RoboDK station: Yuktii_Robotic_Car_Painting_Cell.rdk

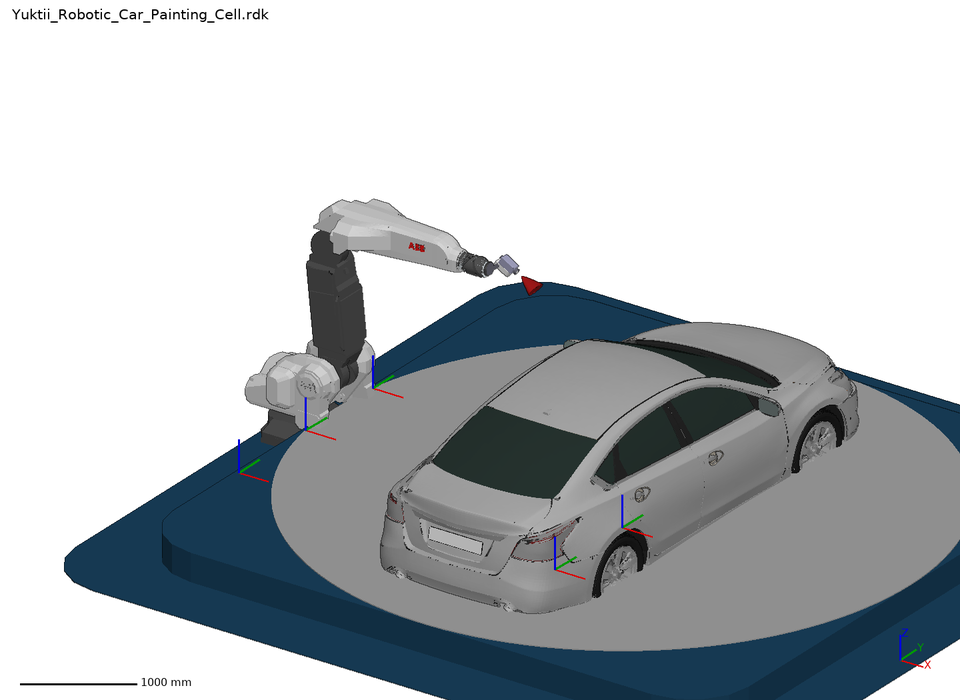
[picture v0: the station drawn from its stored meshes, robots at their saved joint values, targets as dots, program paths as lines]
Station Yuktii_Robotic_Car_Painting_Cell (saved by RoboDK 6.1.1). Poses are relative to the parent item; angles as X-Y-Z fixed-axis rotations.
  - frame ABB IRB 5400-22 Base at (0, 1000, 0) mm
    - robot ABB IRB 5400-22: 6 axes, payload 25 kg, reach 2829 mm, repeatability 0.15 mm, weight 1060 kg
        modified DH rows (alpha deg, a mm, theta deg, d mm): 0, 0, 0, 660; -90, 300, -90, 0; 0, 1200, 0, 0; -90, 213, -90, 1408.298; 35, 0, 0, 79.169; -70, 0, 180, 79.169
        base shift (0, 0, 0) mm, rotated rx 0 ry 0 rz 90 deg
        joint limits [-150, -65, -70, -720, -720, -720] to [150, 150, 70, 720, 720, 720]; home [0, 0, 0, 0, 0, 0]; saved at [-90, 0, 0, -0.001, 0.001, 0.001]
      - tool Generic Paint Sprayer, TCP at (50, 0, 450) mm, rotated rx 0 ry 30 rz 0 deg, size 277.6 x 203.2 x 501.7 mm
    - frame Painting Cell Frame at (0, 0, 0) mm
      - target Home (Cartesian target) at (2370, 0, 2023) mm, rotated rx -180 ry 60 rz -180 deg; joints [-90, 0, 0, 0, 0, 0] of ABB IRB 5400-22
        - target Home (Cartesian target) at (2370, 0, 2023) mm, rotated rx -180 ry 60 rz -180 deg; joints [-90, 0, 0, 0, 0, 0] of ABB IRB 5400-22
      - target Paint_Side_P01 (Cartesian target) at (2687.55, 277.64, 1440.42) mm, rotated rx -179.95 ry 58.29 rz -173.94 deg; joints [-85.31, 17.38, 3.62, 71.65, -55.76, -34.2] of ABB IRB 5400-22
      - target Paint_Side_P02 (Cartesian target) at (2657.17, 535.96, 1322.05) mm, rotated rx 179.9 ry 54.95 rz -168.86 deg; joints [-79.713, 18.918, 5.006, 71.33, -54.978, -34.463] of ABB IRB 5400-22
      - target Paint_Side_P03 (Cartesian target) at (2586.47, 830.84, 1163.47) mm, rotated rx 179.79 ry 50.46 rz -162.52 deg; joints [-73.303, 21.155, 6.646, 70.242, -53.863, -34.183] of ABB IRB 5400-22
      - target Paint_Side_P04 (Cartesian target) at (2523.64, 1053.32, 1068.21) mm, rotated rx 179.74 ry 48.21 rz -157.7 deg; joints [-68.45, 23.41, 6.64, 70.24, -53.86, -34.18] of ABB IRB 5400-22
      - target Paint_Side_P05 (Cartesian target) at (2478.28, 1238.02, 1045.31) mm, rotated rx 179.76 ry 48.45 rz -153.8 deg; joints [-64.55, 25.42, 4.99, 71.3, -54.96, -34.45] of ABB IRB 5400-22
      - target Paint_Side_P06 (Cartesian target) at (2451.93, 1495.48, 1004.92) mm, rotated rx 179.78 ry 49.69 rz -148.94 deg; joints [-59.68, 30.78, -0.3, 73.58, -57.34, -34.99] of ABB IRB 5400-22
      - target Paint_Side_P07 (Cartesian target) at (2459.02, 1865.41, 979.47) mm, rotated rx 179.83 ry 53.14 rz -143.1 deg; joints [-53.79, 41.5, -13.94, 74.57, -58.3, -35.26] of ABB IRB 5400-22
      - target Paint_Side_P08 (Cartesian target) at (2374.12, 1800.72, 860.49) mm, rotated rx 179.76 ry 48.46 rz -143.15 deg; joints [-53.84, 38.265, -5.941, 74.644, -58.451, -35.237] of ABB IRB 5400-22
      - target Paint_Side_P09 (Cartesian target) at (2351.62, 1976.72, 689.21) mm, rotated rx 179.72 ry 46.57 rz -140.3 deg; joints [-50.934, 45.88, -11.622, 74.742, -58.517, -35.278] of ABB IRB 5400-22
      - target Paint_Side_P10 (Cartesian target) at (2340.73, 2028.43, 516.1) mm, rotated rx 179.83 ry 43.58 rz -139.36 deg; joints [-48.072, 50.81, -13.693, -74.012, 58.304, 35.166] of ABB IRB 5400-22
      - target Paint_Side_P11 (Cartesian target) at (2319.85, 2100.8, 404.53) mm, rotated rx 176.79 ry 40.89 rz -141.32 deg; joints [-46.78, 54.89, -17.15, -68.32, 54.72, 34.95] of ABB IRB 5400-22
      - target Paint_Side_P12 (Cartesian target) at (2319.85, 2100.8, 404.53) mm, rotated rx 176.79 ry 40.89 rz -141.32 deg; joints [-48.695, 54.861, -16.957, 73.672, -54.894, -34.206] of ABB IRB 5400-22
      - target Paint_Side_P13 (Cartesian target) at (2357.01, 1967.98, 472.25) mm, rotated rx 176.8 ry 40.88 rz -143.6 deg; joints [-51.025, 50.456, -12.297, 74.028, -55.343, -34.246] of ABB IRB 5400-22
      - target Paint_Side_P14 (Cartesian target) at (2329.44, 1880.14, 669.1) mm, rotated rx 176.66 ry 43.13 rz -144.6 deg; joints [-52.014, 42.506, -6.735, 73.71, -55.102, -34.119] of ABB IRB 5400-22
      - target Paint_Side_P15 (Cartesian target) at (2356.38, 1841.89, 779.16) mm, rotated rx 176.49 ry 45.47 rz -145.61 deg; joints [-52.91, 40.16, -6.73, 73.71, -55.1, -34.11] of ABB IRB 5400-22
      - target Paint_Side_P16 (Cartesian target) at (2375.75, 1666.69, 808.98) mm, rotated rx 176.57 ry 44.12 rz -148.47 deg; joints [-55.911, 35.511, -1.417, 72.415, -53.828, -33.754] of ABB IRB 5400-22
      - target Paint_Side_P17 (Cartesian target) at (2358.71, 1489.22, 826.96) mm, rotated rx 176.71 ry 41.64 rz -151.09 deg; joints [-58.74, 30.11, 4.7, 69.11, -50.54, -32.85] of ABB IRB 5400-22
      - target Paint_Side_P18 (Cartesian target) at (2352.69, 1267.22, 769.5) mm, rotated rx 176.97 ry 36.54 rz -154.8 deg; joints [-62.721, 26.199, 10.485, 62.639, -44.318, -30.826] of ABB IRB 5400-22
      - target Paint_Side_P19 (Cartesian target) at (2339.07, 1164.01, 639.71) mm, rotated rx 177.2 ry 31.03 rz -156.46 deg; joints [-64.56, 26.76, 13.09, 57.4, -39.55, -28.91] of ABB IRB 5400-22
      - target Paint_Side_P20 (Cartesian target) at (2351.97, 1121.3, 477.66) mm, rotated rx 177.35 ry 27.01 rz -157.36 deg; joints [-65.53, 30.78, 13.09, 57.4, -39.55, -28.91] of ABB IRB 5400-22
      - target Paint_Side_P21 (Cartesian target) at (2354.18, 1035.31, 389.95) mm, rotated rx 111.95 ry -49.41 rz 97.65 deg; joints [-61.65, 33.04, 15.16, 173.91, -34.68, -354.54] of ABB IRB 5400-22
      - target Paint_Side_P22 (Cartesian target) at (2300.58, 869.96, 414.39) mm, rotated rx 111.93 ry -49.41 rz 94.75 deg; joints [-64.515, 28.088, 21.499, 170.665, -33.02, -351.904] of ABB IRB 5400-22
      - target Paint_Side_P23 (Cartesian target) at (2314.38, 611.77, 405.59) mm, rotated rx 112.89 ry -49.17 rz 88.15 deg; joints [-70.296, 25.908, 24.902, 169.511, -32.465, -350.855] of ABB IRB 5400-22
      - target Paint_Side_P24 (Cartesian target) at (2342.88, 284.67, 414.82) mm, rotated rx 112.88 ry -49.17 rz 80.3 deg; joints [-78.104, 24.346, 26.702, 169.017, -32.228, -350.379] of ABB IRB 5400-22
      - target Paint_Side_P25 (Cartesian target) at (2359.9, -36.58, 415.09) mm, rotated rx 112.87 ry -49.18 rz 72.49 deg; joints [-85.92, 24.34, 26.7, 169.01, -32.22, -350.37] of ABB IRB 5400-22
      - target Paint_Side_P26 (Cartesian target) at (2326.94, -394.75, 415.09) mm, rotated rx 112.87 ry -49.18 rz 63.75 deg; joints [-94.66, 24.34, 26.7, 169.01, -32.22, -350.37] of ABB IRB 5400-22
      - target Paint_Side_P27 (Cartesian target) at (2252.21, -705.72, 415.09) mm, rotated rx 112.87 ry -49.18 rz 55.98 deg; joints [-102.43, 24.34, 26.7, 169.01, -32.22, -350.37] of ABB IRB 5400-22
      - target Paint_Side_P28 (Cartesian target) at (2279.45, -959.44, 413.25) mm, rotated rx 112.85 ry -49.19 rz 50.17 deg; joints [-107.938, 28.675, 20.449, 174.163, -34.94, -354.053] of ABB IRB 5400-22
      - target Paint_Side_P29 (Cartesian target) at (2329.77, -987.72, 580.14) mm, rotated rx 106.08 ry -50.73 rz 55.16 deg; joints [-108.194, 26.054, 18.009, 175.068, -35.38, -354.858] of ABB IRB 5400-22
      - target Paint_Side_P30 (Cartesian target) at (2366.74, -1005.47, 624.94) mm, rotated rx 104.07 ry -51.08 rz 56.67 deg; joints [-108.306, 26.506, 15.801, 175.982, -35.848, -355.652] of ABB IRB 5400-22
      - target Paint_Side_P31 (Cartesian target) at (2341.49, -1086.77, 693.07) mm, rotated rx 101.34 ry -51.52 rz 56.91 deg; joints [-110.203, 25.189, 15.244, 176.226, -35.966, -355.862] of ABB IRB 5400-22
      - target Paint_Side_P32 (Cartesian target) at (2350.5, -1289.69, 809.61) mm, rotated rx 96.38 ry -52.11 rz 56.93 deg; joints [-114.207, 26.687, 9.223, 179.177, -37.505, -358.342] of ABB IRB 5400-22
      - target Paint_Side_P33 (Cartesian target) at (2338.83, -1380.36, 813.26) mm, rotated rx 96.14 ry -52.14 rz 55.32 deg; joints [-116.05, 28.1, 7.13, 180.3, -38.1, -359.26] of ABB IRB 5400-22
      - target Paint_Side_P34 (Cartesian target) at (2313.09, -1640.06, 805.87) mm, rotated rx 96.12 ry -52.15 rz 50.51 deg; joints [-120.978, 33.486, -0.37, 184.719, -40.559, -362.788] of ABB IRB 5400-22
      - target Paint_Side_P35 (Cartesian target) at (2385.33, -1800.15, 689.63) mm, rotated rx 99.75 ry -51.77 rz 45.91 deg; joints [-122.82, 42.83, -10.73, 191.42, -44.54, -367.93] of ABB IRB 5400-22
      - target Paint_Side_P36 (Cartesian target) at (2352.14, -1838.69, 532.96) mm, rotated rx 104.98 ry -51 rz 40.85 deg; joints [-123.79, 46.18, -10.73, 191.42, -44.54, -367.93] of ABB IRB 5400-22
      - target Paint_Side_P37 (Cartesian target) at (2383.84, -1926.08, 389.53) mm, rotated rx 109 ry -50.23 rz 36.81 deg; joints [-124.76, 53.4, -17.69, 196.12, -47.53, -371.4] of ABB IRB 5400-22
      - target Paint_Side_P38 (Cartesian target) at (2362.81, -2185.89, 442.85) mm, rotated rx 106.5 ry -50.73 rz 34.86 deg; joints [-128.68, 60.25, -31.28, 205.41, -53.93, -377.94] of ABB IRB 5400-22
      - target Paint_Side_P39 (Cartesian target) at (2368.83, -2190.72, 613.31) mm, rotated rx 101.33 ry -51.57 rz 38.89 deg; joints [-128.68, 56.9, -31.28, 205.41, -53.93, -377.94] of ABB IRB 5400-22
      - target Paint_Side_P40 (Cartesian target) at (2364.19, -2186.99, 852.08) mm, rotated rx 93.82 ry -52.34 rz 44.81 deg; joints [-128.68, 52.21, -31.28, 205.41, -53.93, -377.94] of ABB IRB 5400-22
      - target Paint_Side_P41 (Cartesian target) at (2429.25, -2245.53, 801.72) mm, rotated rx 95.27 ry -52.23 rz 43.67 deg; joints [-128.69, 58.91, -40.91, 211.91, -58.84, -382.23] of ABB IRB 5400-22
      - target Paint_Side_P42 (Cartesian target) at (2402.83, -2072.83, 809.3) mm, rotated rx 95.26 ry -52.24 rz 45.66 deg; joints [-126.674, 50.089, -26.385, 202.057, -51.536, -375.626] of ABB IRB 5400-22
      - target Paint_Side_P43 (Cartesian target) at (2397.72, -2068.76, 904.03) mm, rotated rx 92.18 ry -52.45 rz 48.11 deg; joints [-126.67, 48.19, -26.38, 202.05, -51.53, -375.62] of ABB IRB 5400-22
      - target Paint_Side_P44 (Cartesian target) at (2404.71, -1939.77, 930.5) mm, rotated rx 91.34 ry -52.5 rz 50.69 deg; joints [-124.73, 43.5, -19.74, 197.5, -48.43, -372.39] of ABB IRB 5400-22
      - target Paint_Side_P45 (Cartesian target) at (2424.76, -1763.9, 1025.75) mm, rotated rx 88.05 ry -52.62 rz 56.18 deg; joints [-121.803, 37.363, -13.341, 193.148, -45.618, -369.204] of ABB IRB 5400-22
      - target Paint_Side_P46 (Cartesian target) at (2501.66, -1816.71, 1075.26) mm, rotated rx 86.44 ry -52.65 rz 57.5 deg; joints [-121.814, 41.601, -21.433, 198.65, -49.191, -373.214] of ABB IRB 5400-22
      - target Paint_Side_P47 (Cartesian target) at (2521.68, -2035.45, 1120.54) mm, rotated rx 85.17 ry -52.65 rz 55.56 deg; joints [-124.802, 50.228, -36.673, 209.055, -56.613, -380.366] of ABB IRB 5400-22
      - target Paint_Side_P48 (Cartesian target) at (2491.9, -2224.63, 1126.16) mm, rotated rx 85.14 ry -52.65 rz 52.72 deg; joints [-127.67, 58.19, -50.18, 218.04, -63.79, -386.02] of ABB IRB 5400-22
      - target Paint_Side_P49 (Cartesian target) at (2637.88, -1982.32, 1160.05) mm, rotated rx 84.01 ry -52.64 rz 58.46 deg; joints [-122.825, 54.406, -44.865, 214.527, -60.901, -383.866] of ABB IRB 5400-22
      - target Paint_Side_P50 (Cartesian target) at (2582.23, -1809.13, 1242.07) mm, rotated rx 81.02 ry -52.57 rz 62.79 deg; joints [-120.85, 43.5, -29.72, 204.31, -53.12, -377.16] of ABB IRB 5400-22
      - target Paint_Side_P51 (Cartesian target) at (2618.31, -1589.81, 1315.52) mm, rotated rx 74.52 ry -52.89 rz 74.75 deg; joints [-117.93, 36.81, -20.97, 188.74, -39.61, -370.49] of ABB IRB 5400-22
      - target Paint_Side_P52 (Cartesian target) at (2623.91, -1459.92, 1331.56) mm, rotated rx 73.67 ry -52.77 rz 77.67 deg; joints [-115.766, 33.391, -16.372, 184.597, -37.067, -367.591] of ABB IRB 5400-22
      - target Paint_Side_P53 (Cartesian target) at (2616.77, -1306.34, 1411.32) mm, rotated rx 70.58 ry -52.28 rz 82.78 deg; joints [-113.193, 28.706, -12.08, 180.64, -34.713, -364.793] of ABB IRB 5400-22
      - target Paint_Side_P54 (Cartesian target) at (2683.21, -1167.98, 1441.11) mm, rotated rx 69.63 ry -52.12 rz 86.54 deg; joints [-110.175, 28.59, -12.841, 181.347, -35.125, -365.292] of ABB IRB 5400-22
      - target Paint_Side_P55 (Cartesian target) at (2649.23, -855.94, 1495.04) mm, rotated rx 66.81 ry -51.55 rz 94.56 deg; joints [-104.557, 21.072, -4.174, 173.152, -30.436, -359.425] of ABB IRB 5400-22
      - target Paint_Side_P56 (Cartesian target) at (2666.88, -565.19, 1525.15) mm, rotated rx 65.33 ry -51.24 rz 101.73 deg; joints [-98.61, 18.05, -1.14, 170.22, -28.81, -357.3] of ABB IRB 5400-22
      - target Paint_Side_P57 (Cartesian target) at (2662.07, -286.65, 1542.5) mm, rotated rx 64.33 ry -51 rz 108.4 deg; joints [-92.785, 15.593, 1.463, 167.684, -27.43, -355.464] of ABB IRB 5400-22
      - target Paint_Side_P58 (Cartesian target) at (2643.19, -58.71, 1533.21) mm, rotated rx 64.32 ry -51 rz 113.33 deg; joints [-87.918, 14.046, 3.678, 165.507, -26.262, -353.885] of ABB IRB 5400-22
      - target Paint_Side_P59 (Cartesian target) at (2643.6, 168.06, 1475.48) mm, rotated rx 66.28 ry -51.45 rz 116.71 deg; joints [-83.035, 14.713, 4.605, 164.582, -25.771, -353.214] of ABB IRB 5400-22
      - target Home (Cartesian target) at (2370, 0, 2023) mm, rotated rx -180 ry 60 rz 180 deg; joints [-90, 0, 0, -0.001, 0.001, 0] of ABB IRB 5400-22
      - target Target 64 (Cartesian target) at (2431.56, 1366.3, 1005.74) mm, rotated rx 179.72 ry 47.83 rz -151.03 deg; joints [-61.758, 26.931, 4.296, 71.642, -55.315, -34.517] of ABB IRB 5400-22
      - target Target 65 (Cartesian target) at (2421.45, 1107.77, 1017.39) mm, rotated rx 179.66 ry 44.84 rz -155.81 deg; joints [-66.537, 20.959, 10.51, 66.628, -50.22, -33.159] of ABB IRB 5400-22
      - target Target 66 (Cartesian target) at (2437.7, 946.12, 934.72) mm, rotated rx -171.38 ry 35.85 rz -163.72 deg; joints [-66.53, 20.95, 10.5, 66.62, -34.95, -48.93] of ABB IRB 5400-22
      - target Target 67 (Cartesian target) at (2455.17, 839.85, 965.83) mm, rotated rx -149.37 ry 33.2 rz -154.75 deg; joints [-66.53, 20.95, 10.5, 66.62, -34.95, -67.57] of ABB IRB 5400-22
      - target Target 68 (Cartesian target) at (2281.53, 854.15, 1189.47) mm, rotated rx -149.37 ry 33.21 rz -156.42 deg; joints [-63.59, 10.87, 13.54, 58.38, -21.49, -68.41] of ABB IRB 5400-22
      - target Target 69 (Cartesian target) at (2222.52, 748.18, 1108.21) mm, rotated rx -149.07 ry 23.15 rz -166.11 deg; joints [-63.59, 10.87, 13.54, 58.37, -6.99, -76.89] of ABB IRB 5400-22
      - target Target 70 (Cartesian target) at (2314.29, 671.58, 1031.07) mm, rotated rx -174.66 ry 26.9 rz 179.32 deg; joints [-69.41, 12.02, 14.02, 61.4, -11.65, -53.59] of ABB IRB 5400-22
      - target Target 71 (Cartesian target) at (2348.53, 655.22, 1084.89) mm, rotated rx -157.59 ry 30.49 rz -164.86 deg; joints [-69.41, 12.02, 14.02, 44.27, -11.65, -53.59] of ABB IRB 5400-22
      - target Target 72 (Cartesian target) at (2418.39, 483.96, 1040.28) mm, rotated rx -179 ry 31.42 rz 179.44 deg; joints [-76.21, 12.69, 14.02, 44.27, -11.65, -34.95] of ABB IRB 5400-22
      - target Target 73 (Cartesian target) at (2433.89, 322.66, 1024.16) mm, rotated rx -178.61 ry 30.12 rz 175.75 deg; joints [-79.63, 12.635, 13.993, 28.227, -0.687, -26.026] of ABB IRB 5400-22
      - target Target 74 (Cartesian target) at (2450.35, -154.11, 1024.41) mm, rotated rx -178.62 ry 30.13 rz 164.59 deg; joints [-90.78, 12.63, 13.99, 28.22, -0.68, -26.02] of ABB IRB 5400-22
      - target Target 75 (Cartesian target) at (2403.68, -533.92, 1101.06) mm, rotated rx -179.62 ry 33.41 rz 155.34 deg; joints [-100.12, 11.36, 13.92, 47.59, -14.17, -36.57] of ABB IRB 5400-22
      - target Target 76 (Cartesian target) at (2465.14, -650.21, 1055.69) mm, rotated rx -131.01 ry 24.44 rz -156.77 deg; joints [-103.4, 15.42, 13.83, 11.65, -26.09, -42.28] of ABB IRB 5400-22
      - target Target 77 (Cartesian target) at (2445.74, -924.66, 1070.36) mm, rotated rx -129.64 ry 26.09 rz -161.04 deg; joints [-109.805, 18.069, 10.791, 17.454, -31.485, -45.09] of ABB IRB 5400-22
      - target Target 78 (Cartesian target) at (2460.91, -1184.92, 1107) mm, rotated rx -127.19 ry 28.8 rz -163.21 deg; joints [-115.43, 22.74, 4.69, 23.29, -37.86, -47.32] of ABB IRB 5400-22
      - target Target 79 (Cartesian target) at (2442.56, -1519.43, 1130.02) mm, rotated rx -124.71 ry 31.02 rz -166.45 deg; joints [-122.1, 29.121, -3.711, 25.815, -41.925, -47.576] of ABB IRB 5400-22
      - target Target 80 (Cartesian target) at (2573.73, -1565.02, 1176.52) mm, rotated rx -122.14 ry 33.12 rz -163.1 deg; joints [-121.84, 35.09, -12.99, 25.26, -43.26, -46.09] of ABB IRB 5400-22
      - target Target 81 (Cartesian target) at (2490.66, -1694.09, 1176.52) mm, rotated rx -122.14 ry 33.12 rz -166.02 deg; joints [-124.76, 35.09, -12.99, 25.26, -43.26, -46.09] of ABB IRB 5400-22
      - target Target 82 (Cartesian target) at (2506.42, -1705.03, 1062.97) mm, rotated rx -124.25 ry 31.52 rz -167.15 deg; joints [-124.76, 37.48, -12.99, 25.26, -43.26, -46.09] of ABB IRB 5400-22
      - target Target 83 (Cartesian target) at (2447.26, -1788.9, 1062.97) mm, rotated rx -124.25 ry 31.52 rz -169.09 deg; joints [-126.7, 37.48, -12.99, 25.26, -43.26, -46.09] of ABB IRB 5400-22
      - target Target 84 (Cartesian target) at (2436.51, -1757.57, 963.26) mm, rotated rx -126.53 ry 29.7 rz -170.25 deg; joints [-126.265, 37.632, -10.258, 25.738, -43.152, -46.635] of ABB IRB 5400-22
      - target Target 85 (Cartesian target) at (2455.15, -1486.92, 1079.17) mm, rotated rx -108.62 ry 13.32 rz -151.02 deg; joints [-122.27, 29.83, -2.45, 6.99, -44.27, -53.59] of ABB IRB 5400-22
      - target Target 86 (Cartesian target) at (2383.23, -1251.24, 985.09) mm, rotated rx 137.84 ry 45.33 rz 149.2 deg; joints [-127.093, 29.212, 4.635, 62.346, -71.879, 16.542] of ABB IRB 5400-22
      - target Target 87 (Cartesian target) at (2389.27, -903.36, 973.08) mm, rotated rx 136.67 ry 40.82 rz 160.1 deg; joints [-121.56, 24.75, 9.87, 54.4, -70.28, 23.75] of ABB IRB 5400-22
      - target Target 88 (Cartesian target) at (2356.03, -724.5, 1025.32) mm, rotated rx 136.02 ry 38.81 rz 167.16 deg; joints [-119.008, 21.071, 11.864, 47.567, -68.887, 30.048] of ABB IRB 5400-22
      - target Target 89 (Cartesian target) at (2379.15, -397.54, 973.43) mm, rotated rx 134.16 ry 33.87 rz 178.02 deg; joints [-112.26, 21.4, 12.24, 40.3, -67.78, 37.13] of ABB IRB 5400-22
      - target Target 90 (Cartesian target) at (2365.39, -354.45, 922.39) mm, rotated rx 132.55 ry 30.09 rz -178.82 deg; joints [-111.726, 22.838, 11.574, 35.485, -67.33, 42.068] of ABB IRB 5400-22
      - target Target 91 (Cartesian target) at (2377.11, -152.88, 925.3) mm, rotated rx 132.01 ry 28.94 rz -172.71 deg; joints [-107.078, 22.996, 10.964, 33.204, -67.266, 44.598] of ABB IRB 5400-22
      - target Target 93 (Cartesian target) at (2365.62, 454.26, 908.58) mm, rotated rx -180 ry 29.04 rz -169.13 deg; joints [-79.13, 12.02, 18.94, 0, 0, 0] of ABB IRB 5400-22
      - target Target 93 (Cartesian target) at (2307.39, 692.25, 908.9) mm, rotated rx -180 ry 29.05 rz -163.3 deg; joints [-73.3, 12.02, 18.93, 0, 0, 0] of ABB IRB 5400-22
      - target Target 94 (Cartesian target) at (2321.31, 696.8, 661.14) mm, rotated rx 179.99 ry 22.35 rz -163.31 deg; joints [-73.29, 18.72, 18.93, -0.01, 0.02, 0.01] of ABB IRB 5400-22
      - target Target 96 (Cartesian target) at (2265.55, 985.02, 820.27) mm, rotated rx 179.99 ry 29.71 rz -156.52 deg; joints [-65.754, 16.526, 17.771, -34.157, 22.81, 19.698] of ABB IRB 5400-22
      - target Target 96 (Cartesian target) at (2355.77, 1024.1, 856.74) mm, rotated rx 179.89 ry 35.33 rz -156.57 deg; joints [-65.504, 19.848, 14.513, -52.037, 36.976, 28.267] of ABB IRB 5400-22
      - target Target 97 (Cartesian target) at (2297.33, 1237.75, 742.18) mm, rotated rx 179.94 ry 33.8 rz -151.73 deg; joints [-60.656, 24.16, 13.203, -55.596, 40.098, 29.701] of ABB IRB 5400-22
      - target Target 99 (Cartesian target) at (2334.09, -1564.72, 911.12) mm, rotated rx 179.66 ry 44.54 rz 145.94 deg; joints [-122.78, 29.44, 3.24, -68.04, 51.94, 33.9] of ABB IRB 5400-22
      - target Target 99 (Cartesian target) at (2383.08, -1922.61, 792.43) mm, rotated rx 129.8 ry 40.18 rz 114.6 deg; joints [-131.6, 45.51, -12.13, -71.68, 58.25, 72.23] of ABB IRB 5400-22
      - target Target 100 (Cartesian target) at (2320.47, -1611.26, 821.25) mm, rotated rx 131.5 ry 37.1 rz 123.46 deg; joints [-128.622, 34.639, 2.593, -77.933, 59.044, 77.036] of ABB IRB 5400-22
      - target Target 101 (Cartesian target) at (2345.57, -1090.33, 826.64) mm, rotated rx 133.32 ry 31.79 rz 139.56 deg; joints [-120.514, 24.999, 14.295, -81.52, 53.807, 82.959] of ABB IRB 5400-22
      - target Target 102 (Cartesian target) at (2357.6, -322.96, 677.83) mm, rotated rx 134.67 ry 19.27 rz 165.08 deg; joints [-105.77, 21.651, 21.251, -84.321, 41.712, 92.046] of ABB IRB 5400-22
      - target Target 103 (Cartesian target) at (2336.63, 1100.19, 539.42) mm, rotated rx -169.54 ry 29.49 rz -173.27 deg; joints [-57.41, 31.45, 10.05, -33.99, 55.09, -1.39] of ABB IRB 5400-22
      - target Target 104 (Cartesian target) at (2301.03, -953.45, 610.69) mm, rotated rx 143.59 ry 28.63 rz 126.15 deg; joints [-112.14, 23.41, 22.34, -54.77, 58.25, 53.59] of ABB IRB 5400-22
      - target Target 105 (Cartesian target) at (2332.17, -895.94, 508.39) mm, rotated rx 131.34 ry 21.29 rz 122.4 deg; joints [-112.14, 27.43, 22.34, -54.77, 58.24, 67.57] of ABB IRB 5400-22
      - target Target 106 (Cartesian target) at (2329.78, 1096.4, 434.09) mm, rotated rx -168.24 ry 27.08 rz -172.64 deg; joints [-57.4, 34.13, 10.04, -33.99, 55.09, -1.38] of ABB IRB 5400-22
      - target Home (Cartesian target) at (2370, 0, 2023) mm, rotated rx -180 ry 60 rz -180 deg; joints [-90, 0, 0, 0, 0, 0] of ABB IRB 5400-22
      - target New_Side1 (Cartesian target) at (2658.8, 275.75, 1524.52) mm, rotated rx -179.85 ry 60.31 rz -173.84 deg; joints [-85.3, 15.37, 3.61, 71.65, -55.76, -34.2] of ABB IRB 5400-22
      - target Target 108 (Cartesian target) at (2664.22, 523.99, 1523.09) mm, rotated rx -179.82 ry 60.98 rz -168.61 deg; joints [-80.075, 17.43, 1.429, 72.616, -56.756, -34.445] of ABB IRB 5400-22
      - target Target 109 (Cartesian target) at (2665.93, 762.89, 1510.03) mm, rotated rx -179.81 ry 61.52 rz -163.77 deg; joints [-75.205, 20.33, -1.486, 73.532, -57.694, -34.668] of ABB IRB 5400-22
      - target Target 110 (Cartesian target) at (2659.82, 1167.43, 1438.23) mm, rotated rx -179.83 ry 61.51 rz -156.05 deg; joints [-67.415, 27.34, -7.983, 74.44, -58.603, -34.91] of ABB IRB 5400-22
      - target Target 111 (Cartesian target) at (2634.53, 1372.82, 1374.32) mm, rotated rx -179.9 ry 60.79 rz -152.28 deg; joints [-63.559, 31.151, -11.105, 74.432, -58.556, -34.922] of ABB IRB 5400-22
      - target Target 112 (Cartesian target) at (2613.56, 1565.5, 1326.63) mm, rotated rx -156.73 ry 55.5 rz -141.8 deg; joints [-57.009, 36.126, -17.739, 72.955, -48.745, -56.751] of ABB IRB 5400-22
      - target Target 113 (Cartesian target) at (2569.84, 1720.18, 1273.47) mm, rotated rx -156.83 ry 54.94 rz -138.73 deg; joints [-54.23, 38.988, -20.195, 72.171, -48.363, -56.199] of ABB IRB 5400-22
      - target Target 114 (Cartesian target) at (2584.39, 1876.48, 1194.72) mm, rotated rx -130.83 ry 49.71 rz -130.74 deg; joints [-48.997, 49.602, -32.053, 80.685, -47.963, -85.459] of ABB IRB 5400-22
      - target Target 115 (Cartesian target) at (2561.17, 2039.05, 1143.93) mm, rotated rx -130.84 ry 49.71 rz -126.9 deg; joints [-46.823, 54.832, -38.834, 75.333, -44.25, -82.66] of ABB IRB 5400-22
      - target Target 116 (Cartesian target) at (2560.42, 2235.82, 1117.58) mm, rotated rx -130.52 ry 50.72 rz -122.04 deg; joints [-44.699, 64.532, -54.336, 60.957, -33.248, -75.821] of ABB IRB 5400-22
      - target Target 117 (Cartesian target) at (2472.08, 1830.68, 1089.48) mm, rotated rx -131.27 ry 45.32 rz -133.48 deg; joints [-47.68, 44.84, -21.46, 88.72, -52.51, -90.54] of ABB IRB 5400-22
      - target Target 118 (Cartesian target) at (2481.64, 1840.12, 992.4) mm, rotated rx -131.47 ry 43.32 rz -133.61 deg; joints [-47.67, 46.85, -21.46, 88.72, -52.51, -90.54] of ABB IRB 5400-22
      - target Target 119 (Cartesian target) at (2403.75, 1952.84, 974.82) mm, rotated rx -131.49 ry 43.1 rz -131.1 deg; joints [-45.15, 47.52, -21.91, 88.72, -52.51, -90.54] of ABB IRB 5400-22
      - target Target 120 (Cartesian target) at (2386.21, 2042.31, 939.94) mm, rotated rx -118.24 ry 38.52 rz -123.55 deg; joints [-43.2, 52.21, -26.67, 84.98, -50.64, -100.19] of ABB IRB 5400-22
      - target Target 121 (Cartesian target) at (2451.41, 2090.3, 884.4) mm, rotated rx -118.24 ry 38.52 rz -121.61 deg; joints [-43.82, 57.066, -32.806, 78.784, -47.107, -96.687] of ABB IRB 5400-22
      - target Target 122 (Cartesian target) at (2455.32, 2094.41, 790.53) mm, rotated rx -118.74 ry 36.71 rz -121.91 deg; joints [-43.82, 58.91, -32.8, 78.78, -47.1, -96.68] of ABB IRB 5400-22
      - target Target 123 (Cartesian target) at (2455.32, 2094.41, 790.53) mm, rotated rx -118.74 ry 36.71 rz -121.91 deg; joints [-43.82, 58.91, -32.8, 78.78, -47.1, -96.68] of ABB IRB 5400-22
      - target Target 124 (Cartesian target) at (2404.28, 2248.71, 785.39) mm, rotated rx -105.86 ry 31.76 rz -113.98 deg; joints [-40.99, 65.21, -41.48, 70.02, -41.43, -104.85] of ABB IRB 5400-22
      - target Target 125 (Cartesian target) at (2471.68, 2333.46, 771.99) mm, rotated rx -105.61 ry 32.35 rz -110.71 deg; joints [-41.26, 72.98, -55.01, 51.48, -28.89, -95.09] of ABB IRB 5400-22
      - target Target 126 (Cartesian target) at (2420.97, 2346.66, 641.9) mm, rotated rx -106.69 ry 29.85 rz -111.27 deg; joints [-40.388, 73.008, -50.637, 57.956, -33.304, -98.515] of ABB IRB 5400-22
      - target Target 127 (Cartesian target) at (2419.04, 2345.11, 536.48) mm, rotated rx -107.43 ry 27.97 rz -111.62 deg; joints [-40.38, 74.98, -50.63, 57.95, -33.3, -98.51] of ABB IRB 5400-22
      - target Target 128 (Cartesian target) at (2416.56, 2342.24, 464.73) mm, rotated rx -107.92 ry 26.7 rz -111.84 deg; joints [-40.38, 76.32, -50.62, 57.95, -33.3, -98.5] of ABB IRB 5400-22
      - target Target 129 (Cartesian target) at (2372.36, 2151.25, 436.56) mm, rotated rx -108.49 ry 24.41 rz -118.69 deg; joints [-41.3, 67.62, -33.69, 79.97, -47.44, -109.64] of ABB IRB 5400-22
      - target Target 130 (Cartesian target) at (2332.85, 1868.98, 420.57) mm, rotated rx -108.74 ry 20.64 rz -131.35 deg; joints [-42.87, 60.25, -19.97, 102.16, -57.85, -121.49] of ABB IRB 5400-22
      - target Target 131 (Cartesian target) at (2362.92, 1786.92, 599.14) mm, rotated rx -108.64 ry 23.66 rz -135.23 deg; joints [-44.065, 55.5, -18.473, 106.546, -59.354, -124.195] of ABB IRB 5400-22
      - target Target 132 (Cartesian target) at (2352.74, 1670.01, 745.54) mm, rotated rx -108.35 ry 24.36 rz -143.99 deg; joints [-44.63, 51.54, -17.35, 119.07, -63.26, -132.98] of ABB IRB 5400-22
      - target Target 133 (Cartesian target) at (2352.74, 1670.01, 745.54) mm, rotated rx -108.35 ry 24.36 rz -143.99 deg; joints [-44.63, 51.54, -17.35, 119.07, -63.26, -132.98] of ABB IRB 5400-22
      - target Target 134 (Cartesian target) at (2336.83, 1664.58, 784.26) mm, rotated rx -108.35 ry 24.36 rz -146.45 deg; joints [-44.2, 51.085, -18.114, 123.264, -64.411, -136.171] of ABB IRB 5400-22
      - target Target 135 (Cartesian target) at (2327.68, 1352.65, 832.3) mm, rotated rx -103.03 ry 1.48 rz -109.02 deg; joints [-54.222, 28.746, 9.244, -28.437, 5.83, -416.904] of ABB IRB 5400-22
      - target Target 136 (Cartesian target) at (2306.29, 1190.11, 834.99) mm, rotated rx -103.59 ry 0.51 rz -109.04 deg; joints [-57.25, 24.08, 15.62, -46.54, 14.38, -405.66] of ABB IRB 5400-22
      - target Target 137 (Cartesian target) at (2334.57, 1071.93, 714.75) mm, rotated rx -105.67 ry -2.13 rz -112.44 deg; joints [-59.663, 25.899, 17.118, -42.65, 12.894, -408.122] of ABB IRB 5400-22
      - target Target 138 (Cartesian target) at (2330.83, 977.71, 595.32) mm, rotated rx -107.81 ry -4.94 rz -115.26 deg; joints [-61.28, 27.482, 18.954, -36.885, 10.544, -411.674] of ABB IRB 5400-22
      - target Target 174 (Cartesian target) at (2370, 0, 2023) mm, rotated rx -180 ry 60 rz -180 deg; joints [-90, 0, 0, 0, 0, 0] of ABB IRB 5400-22
      - target Target 175 (Cartesian target) at (2003.56, 0, 1478.8) mm, rotated rx -180 ry 46.35 rz -180 deg; joints [-90, -16.78, 30.43, 0, 0, 0] of ABB IRB 5400-22
      - target Target 140 (Cartesian target) at (2346.95, 903.39, 372.64) mm, rotated rx 105.05 ry -53.98 rz 91.43 deg; joints [-62.798, 32.643, 18.247, 171.995, -33.643, 20.163] of ABB IRB 5400-22
      - target Target 141 (Cartesian target) at (2342.97, 174.12, 368.94) mm, rotated rx 106.29 ry -53.62 rz 73.14 deg; joints [-79.038, 26.889, 26.977, 168.799, -32.261, 24.129] of ABB IRB 5400-22
      - target Target 142 (Cartesian target) at (2350.11, -835.78, 365.76) mm, rotated rx 105.46 ry -53.86 rz 50.44 deg; joints [-103.37, 32.12, 19.32, 171.49, -33.41, 20.69] of ABB IRB 5400-22
      - target Target 143 (Cartesian target) at (2337.88, -1111.77, 373.69) mm, rotated rx 100.3 ry -27.32 rz 78.87 deg; joints [-114.08, 34.8, 19.32, 123.5, -33.41, 25.63] of ABB IRB 5400-22
      - target Target 145 (Cartesian target) at (2293.54, -1236.73, 723.48) mm, rotated rx 90.92 ry -25.06 rz 80.1 deg; joints [-116.99, 26.09, 19.32, 123.5, -33.41, 25.63] of ABB IRB 5400-22
      - target Target 146 (Cartesian target) at (2289.45, -1364.49, 777.87) mm, rotated rx 89.51 ry -24.66 rz 77.78 deg; joints [-119.341, 27.215, 15.821, 125.411, -33.698, 23.861] of ABB IRB 5400-22
      - target Target 147 (Cartesian target) at (2331.68, -1489.87, 827.19) mm, rotated rx 88.33 ry -24.33 rz 75.77 deg; joints [-120.96, 30.317, 9.647, 128.755, -34.187, 20.613] of ABB IRB 5400-22
      - target Target 148 (Cartesian target) at (2325.53, -1697.75, 857.4) mm, rotated rx 90.71 ry -12.89 rz 74.04 deg; joints [-124.76, 34.8, 3.22, 131.19, -44.16, 13.4] of ABB IRB 5400-22
      - target Target 149 (Cartesian target) at (2344.83, -1796.94, 780.88) mm, rotated rx 92.31 ry -13.4 rz 71.83 deg; joints [-125.99, 39.49, -1.41, 132.9, -44.03, 11.23] of ABB IRB 5400-22
      - target Target 150 (Cartesian target) at (2326.9, -1929.07, 663.98) mm, rotated rx 94.68 ry -14.1 rz 68.63 deg; joints [-128.1, 44.84, -5.96, 134.54, -43.87, 9.06] of ABB IRB 5400-22
      - target Target 151 (Cartesian target) at (2330.1, -2009.3, 463.73) mm, rotated rx 98.67 ry -15.23 rz 66.11 deg; joints [-129.136, 51.704, -10.429, 136.139, -43.668, 6.9] of ABB IRB 5400-22
      - target Target 152 (Cartesian target) at (2324.17, -2004.03, 374.06) mm, rotated rx 100.53 ry -15.71 rz 65.62 deg; joints [-129.13, 53.55, -10.42, 136.13, -43.66, 6.9] of ABB IRB 5400-22
      - target Target 153 (Cartesian target) at (2350.91, -2138.26, 409.75) mm, rotated rx 95.5 ry -11.04 rz 69.58 deg; joints [-131.63, 58.24, -17.66, 125.27, -42.28, 12.86] of ABB IRB 5400-22
      - target Target 154 (Cartesian target) at (2358.16, -2144.71, 578.33) mm, rotated rx 92.34 ry -9.81 rz 70.15 deg; joints [-131.63, 54.89, -17.66, 125.27, -42.28, 12.86] of ABB IRB 5400-22
      - target Target 155 (Cartesian target) at (2351.78, -2034.83, 598.74) mm, rotated rx 92.01 ry -9.71 rz 72.24 deg; joints [-130.35, 50.87, -11.47, 123.69, -43.37, 15.86] of ABB IRB 5400-22
      - target Target 156 (Cartesian target) at (2361.73, -2031.04, 641.31) mm, rotated rx 91.21 ry -9.37 rz 72.51 deg; joints [-130.17, 50.2, -11.81, 123.77, -43.3, 15.68] of ABB IRB 5400-22
      - target Target 157 (Cartesian target) at (2381.46, -2007.86, 641.31) mm, rotated rx 91.21 ry -9.37 rz 73.07 deg; joints [-129.61, 50.2, -11.81, 123.77, -43.3, 15.68] of ABB IRB 5400-22
      - target Target 158 (Cartesian target) at (2371.55, -1954.82, 707.1) mm, rotated rx 89.96 ry -8.85 rz 74.24 deg; joints [-129.052, 47.01, -8.72, 122.993, -43.864, 17.153] of ABB IRB 5400-22
      - target Target 159 (Cartesian target) at (2375.07, -1837.16, 777.79) mm, rotated rx 88.57 ry -8.25 rz 76.8 deg; joints [-127.418, 42.553, -3.828, 121.744, -44.753, 19.458] of ABB IRB 5400-22
      - target Target 160 (Cartesian target) at (2381.93, -1755.68, 825.25) mm, rotated rx 87.62 ry -7.82 rz 78.62 deg; joints [-126.181, 39.789, -1.019, 121.01, -45.257, 20.759] of ABB IRB 5400-22
      - target Target 161 (Cartesian target) at (2414.53, -1737.26, 915.15) mm, rotated rx 85.9 ry -7.01 rz 79.3 deg; joints [-125.47, 38.82, -2.55, 121.42, -44.98, 20.01] of ABB IRB 5400-22
      - target Target 162 (Cartesian target) at (2430.75, -1523.5, 926.8) mm, rotated rx 85.49 ry -6.84 rz 83.96 deg; joints [-122.07, 34.13, 4.33, 119.51, -46.13, 23.25] of ABB IRB 5400-22
      - target Target 163 (Cartesian target) at (2440.67, -1339.39, 956.51) mm, rotated rx 84.74 ry -6.46 rz 88.16 deg; joints [-118.98, 30.11, 9.37, 118.02, -46.96, 25.58] of ABB IRB 5400-22
      - target Target 164 (Cartesian target) at (2475.14, -1166.95, 1009.48) mm, rotated rx 83.54 ry -5.85 rz 92.22 deg; joints [-115.594, 27.22, 11.797, 117.241, -47.321, 26.717] of ABB IRB 5400-22
      - target Target 165 (Cartesian target) at (2541.7, -966.33, 1114.32) mm, rotated rx 81.35 ry -4.68 rz 96.85 deg; joints [-111.17, 24.75, 11.79, 117.24, -47.32, 26.71] of ABB IRB 5400-22
      - target Target 166 (Cartesian target) at (2438.77, -1046.57, 1116.61) mm, rotated rx 127.47 ry 31.35 rz 100.95 deg; joints [-111.17, 19.39, 11.78, 123.5, -62.91, -30.29] of ABB IRB 5400-22
      - target Target 167 (Cartesian target) at (2502.55, -919.8, 1181.69) mm, rotated rx 125.46 ry 32.41 rz 102.81 deg; joints [-108.097, 19.012, 10.424, 123.971, -63.426, -30.24] of ABB IRB 5400-22
      - target Target 168 (Cartesian target) at (2593.39, -572.94, 1327.96) mm, rotated rx 121.36 ry 34.36 rz 108.17 deg; joints [-100.33, 16.71, 9.02, 124.4, -63.89, -30.21] of ABB IRB 5400-22
      - target Target 169 (Cartesian target) at (2593.39, -572.94, 1327.96) mm, rotated rx 121.36 ry 34.36 rz 108.17 deg; joints [-100.33, 16.71, 9.02, 124.4, -63.89, -30.21] of ABB IRB 5400-22
      - target Target 170 (Cartesian target) at (2606.86, -356.08, 1410.12) mm, rotated rx 119.19 ry 35.3 rz 111.63 deg; joints [-95.63, 14.7, 9.02, 124.4, -63.89, -30.21] of ABB IRB 5400-22
      - target Target 171 (Cartesian target) at (2660.01, 12.46, 1498.43) mm, rotated rx 116.04 ry 36.56 rz 117.57 deg; joints [-87.53, 15.37, 5.88, 125.22, -64.73, -30.24] of ABB IRB 5400-22
      - target Target 172 (Cartesian target) at (2657.4, 365.18, 1513.99) mm, rotated rx 115.28 ry 36.85 rz 124.54 deg; joints [-79.958, 16.341, 4.355, 125.548, -65.04, -30.288] of ABB IRB 5400-22
      - target Home (Cartesian target) at (2370, 0, 2023) mm, rotated rx -180 ry 60 rz -180 deg; joints [-90, 0, 0, 0, 0, 0] of ABB IRB 5400-22
      - target Target 175 (Cartesian target) at (2472.08, 1830.68, 1089.48) mm, rotated rx -131.27 ry 45.32 rz -133.48 deg; joints [-47.68, 44.84, -21.46, 88.72, -52.51, -90.54] of ABB IRB 5400-22
      - target Target 176 (Cartesian target) at (2427.86, 1264.35, 1099.18) mm, rotated rx -130.5 ry 36.23 rz -154.16 deg; joints [-53.543, 32.02, -4.416, 109.606, -56.215, -109.469] of ABB IRB 5400-22
      - target Target 177 (Cartesian target) at (2382.88, -673.82, 1025.37) mm, rotated rx -179.04 ry 31.47 rz 152.37 deg; joints [-103.4, 13.36, 13.92, 47.58, -14.16, -36.56] of ABB IRB 5400-22
      - target Target 178 (Cartesian target) at (2295.9, -645.43, 1322.87) mm, rotated rx 178.75 ry 38.01 rz 151.12 deg; joints [-102.66, 4.66, 13.84, 21.49, 3.52, -21.94] of ABB IRB 5400-22
      - target Target 179 (Cartesian target) at (2289.84, -801.89, 1175.32) mm, rotated rx -179.9 ry 34.14 rz 148.27 deg; joints [-106.31, 8.68, 13.84, 21.49, 3.52, -21.94] of ABB IRB 5400-22
      - target Target 180 (Cartesian target) at (2275.94, -840.54, 1175.32) mm, rotated rx -179.9 ry 34.14 rz 147.3 deg; joints [-107.28, 8.68, 13.84, 21.49, 3.52, -21.94] of ABB IRB 5400-22
      - target Target 181 (Cartesian target) at (2192.36, -786.89, 1107.97) mm, rotated rx -179.9 ry 34.14 rz 147.3 deg; joints [-105.797, 5.265, 20.224, -4.848, 20.771, -6.041] of ABB IRB 5400-22
      - target Target 182 (Cartesian target) at (2382.86, -994.11, 973.37) mm, rotated rx 178.01 ry 39.71 rz 144.57 deg; joints [-108.817, 18.689, 12.609, -41.483, 44.688, 16.144] of ABB IRB 5400-22
      - target Target 183 (Cartesian target) at (2400.81, -1006.99, 991.61) mm, rotated rx 177.52 ry 40.97 rz 144.26 deg; joints [-108.962, 19.291, 11.631, -43.669, 46.321, 17.307] of ABB IRB 5400-22
      - target Target 184 (Cartesian target) at (2376.37, -1347.22, 1008.7) mm, rotated rx 145.79 ry 38.45 rz 130.25 deg; joints [-121.27, 24.75, 5.8, -54.81, 42.93, 54.56] of ABB IRB 5400-22
      - target Target 185 (Cartesian target) at (2422.65, -1754.66, 920.86) mm, rotated rx 128.56 ry 37.29 rz 115.93 deg; joints [-128.64, 39.35, -8.65, -60.74, 49.18, 70.09] of ABB IRB 5400-22
      - target Target 186 (Cartesian target) at (2354.37, -1824.66, 835.51) mm, rotated rx 129.7 ry 35.34 rz 115.04 deg; joints [-130.58, 40.29, -7.39, -61.24, 49.21, 70.51] of ABB IRB 5400-22
      - target Target 187 (Cartesian target) at (2377.86, -1153.27, 879.75) mm, rotated rx 132.19 ry 29.42 rz 134.82 deg; joints [-120.75, 25.42, 10.41, -65.41, 42.63, 77.65] of ABB IRB 5400-22
      - target Target 188 (Cartesian target) at (2359.94, -929.24, 826.9) mm, rotated rx 133.34 ry 24.54 rz 142.99 deg; joints [-117.419, 22.585, 14.742, -64.911, 36.511, 80.455] of ABB IRB 5400-22
      - target Target 189 (Cartesian target) at (2391.23, -667.17, 827.39) mm, rotated rx 133.65 ry 22.34 rz 150.99 deg; joints [-112.14, 20.73, 16.41, -64.25, 32.39, 82.07] of ABB IRB 5400-22
      - target Target 190 (Cartesian target) at (2202.62, -831.48, 1034.88) mm, rotated rx 133.65 ry 22.34 rz 150.99 deg; joints [-118.843, 12.15, 18.199, -62.412, 21.357, 86.632] of ABB IRB 5400-22
      - target Target 191 (Cartesian target) at (2109.76, -912.38, 1137.03) mm, rotated rx 133.65 ry 22.34 rz 150.99 deg; joints [-122.36, 8.718, 17.956, -62.764, 16.398, 90.091] of ABB IRB 5400-22
      - target Target 192 (Cartesian target) at (2280.41, -644.54, 1108.05) mm, rotated rx 155.69 ry 31.8 rz 164.39 deg; joints [-111.17, 8.68, 17.95, -58.25, 20.97, 62.91] of ABB IRB 5400-22
      - target Target 193 (Cartesian target) at (2291.01, -605.37, 1108.38) mm, rotated rx 155.69 ry 31.81 rz 165.37 deg; joints [-110.19, 8.67, 17.95, -58.24, 20.96, 62.91] of ABB IRB 5400-22
      - target Target 194 (Cartesian target) at (2368.73, -670.39, 889.33) mm, rotated rx -161.9 ry 27.55 rz -170.95 deg; joints [-106.31, 14.7, 17.95, -67.57, 25.63, 30.29] of ABB IRB 5400-22
      - target Target 195 (Cartesian target) at (2390.69, -115.75, 865.83) mm, rotated rx -164.07 ry 23.28 rz -159.26 deg; joints [-93.654, 12.603, 19.045, -35.861, 2.338, 14.58] of ABB IRB 5400-22
      - target Target 196 (Cartesian target) at (2355.61, 340.8, 891.86) mm, rotated rx 176.44 ry 30.26 rz 172.94 deg; joints [-78.181, 11.623, 20.691, -16.162, 28.516, 5.142] of ABB IRB 5400-22
      - target Target 197 (Cartesian target) at (2340.91, 486.87, 938.41) mm, rotated rx -175.27 ry 39.05 rz 171.84 deg; joints [-70.439, 13.268, 20.61, -39.821, 58.372, 2.503] of ABB IRB 5400-22
      - target Target 198 (Cartesian target) at (2390.18, 1030.97, 973.44) mm, rotated rx -175.27 ry 39.05 rz 171.84 deg; joints [-57.416, 24.788, 4.133, -31.939, 65.368, -10.181] of ABB IRB 5400-22
      - target Target 199 (Cartesian target) at (2421.98, 1792.86, 985.86) mm, rotated rx -173.33 ry 37.83 rz 173.05 deg; joints [-44.166, 50.231, -35.31, -18.806, 69, -32.901] of ABB IRB 5400-22
      - target Target 200 (Cartesian target) at (2431.65, 1968.76, 881.88) mm, rotated rx -170.66 ry 36.26 rz 174.67 deg; joints [-41.902, 61.657, -50.904, -13.725, 68.144, -41.082] of ABB IRB 5400-22
      - target Target 201 (Cartesian target) at (2358.89, 1432.26, 912.73) mm, rotated rx -170.66 ry 36.26 rz 174.67 deg; joints [-48.958, 35.938, -10.401, -25.18, 68.51, -22.557] of ABB IRB 5400-22
      - target Target 202 (Cartesian target) at (2357.62, 1014.78, 861.63) mm, rotated rx -170.66 ry 36.26 rz 174.67 deg; joints [-57.208, 25.701, 6.641, -31.782, 65.111, -11.655] of ABB IRB 5400-22
      - target Target 203 (Cartesian target) at (2353.37, 451.37, 804.48) mm, rotated rx -179.86 ry 36.82 rz 171.57 deg; joints [-72.66, 15.55, 22.8, -44.27, 58.25, 11.65] of ABB IRB 5400-22
      - target Target 204 (Cartesian target) at (2334.74, -1169.14, 724.21) mm, rotated rx -179.32 ry 35.32 rz -178.39 deg; joints [-122.233, 27.53, 11.574, -119.445, 63.194, 66.577] of ABB IRB 5400-22
      - target Target 205 (Cartesian target) at (2350.16, -1037.89, 637.17) mm, rotated rx 178 ry 31.92 rz -176.57 deg; joints [-119.68, 28.1, 13.25, -119.34, 61.38, 68.24] of ABB IRB 5400-22
      - target Target 207 (Cartesian target) at (2353, -10.72, 730.37) mm, rotated rx 173.9 ry 37.05 rz -171.74 deg; joints [-93.095, 14.814, 28.584, -93.88, 60.635, 53.648] of ABB IRB 5400-22
      - target Target 207 (Cartesian target) at (2350.88, 491.32, 683.54) mm, rotated rx -169.01 ry 37.68 rz -168.12 deg; joints [-73.86, 18.05, 26.54, -69.09, 62.77, 20.43] of ABB IRB 5400-22
      - target Target 208 (Cartesian target) at (2325.13, 1002.17, 663.71) mm, rotated rx -169.8 ry 39.7 rz -168.61 deg; joints [-59.767, 25.598, 17.777, -59.826, 69.712, 10.399] of ABB IRB 5400-22
      - target Target 209 (Cartesian target) at (2345, 916.78, 513.76) mm, rotated rx -168.26 ry 36.06 rz -168.23 deg; joints [-61.997, 28.913, 18.7, -61.531, 69.535, 11.732] of ABB IRB 5400-22
      - target Target 210 (Cartesian target) at (2373.7, 432.14, 423.97) mm, rotated rx -168 ry 31.45 rz -168.09 deg; joints [-75.55, 26.09, 25.68, -71.88, 64.23, 21.26] of ABB IRB 5400-22
      - target Target 211 (Cartesian target) at (2346.62, -866.85, 439.55) mm, rotated rx -175.56 ry 21.24 rz -171.45 deg; joints [-114.24, 29.44, 15.94, -106.79, 47.09, 57.55] of ABB IRB 5400-22
      - target Target 212 (Cartesian target) at (2360.24, -1116.55, 456.2) mm, rotated rx -176.21 ry 20.49 rz -171.67 deg; joints [-120.07, 34.13, 7.98, -116.27, 47.48, 65.53] of ABB IRB 5400-22
      - target Home (Cartesian target) at (2370, 0, 2023) mm, rotated rx -180 ry 60 rz -180 deg; joints [-90, 0, 0, 0, 0, 0] of ABB IRB 5400-22
      - target Target 224 (Cartesian target) at (2388.86, 1869.5, 1172.96) mm, rotated rx 176.01 ry 42.73 rz -145.65 deg; joints [-51.94, 36.14, -18.94, 0, 1.97, 1.81] of ABB IRB 5400-22
      - target Target 225 (Cartesian target) at (2208.58, 1826.17, 1215.73) mm, rotated rx 176.14 ry 41.23 rz -144.03 deg; joints [-50.4, 27.43, -8.72, 0, 1.97, 1.81] of ABB IRB 5400-22
      - target Target 226 (Cartesian target) at (2003.14, 1703.87, 1199.13) mm, rotated rx 176.37 ry 38.34 rz -143.08 deg; joints [-49.6, 16.71, 4.89, 0, 1.97, 1.81] of ABB IRB 5400-22
      - target Backside_Half (Cartesian target) at (1816.9, 1523.09, 1167.51) mm, rotated rx 176.52 ry 36.11 rz -143.4 deg; joints [-50.01, 5.33, 18.51, 0, 1.98, 1.82] of ABB IRB 5400-22
      - target Target 215 (Cartesian target) at (1638.76, 1274.29, 1156.33) mm, rotated rx 176.53 ry 36.11 rz -145.71 deg; joints [-51.94, -8.76, 32.7, -3.28, 4.38, 3.61] of ABB IRB 5400-22
      - target Target 216 (Cartesian target) at (1522.9, 1053.07, 1147.52) mm, rotated rx 176.36 ry 37.87 rz -149.34 deg; joints [-54.85, -20.79, 43.19, -6.92, 7.26, 5.48] of ABB IRB 5400-22
      - target Target 217 (Cartesian target) at (1509.52, 969.02, 1180.46) mm, rotated rx 176.17 ry 39.76 rz -151.41 deg; joints [-56.8, -24.81, 45.32, -6.92, 7.26, 5.48] of ABB IRB 5400-22
      - target Target 218 (Cartesian target) at (1305.45, 1074.88, 1153.68) mm, rotated rx 176.07 ry 40.68 rz -144.67 deg; joints [-50, -30.84, 50.43, -6.92, 7.26, 5.48] of ABB IRB 5400-22
      - target Target 219 (Cartesian target) at (1423.96, 1174.33, 1165.62) mm, rotated rx 176.3 ry 38.54 rz -144.52 deg; joints [-50, -21.46, 43.19, -6.91, 7.25, 5.47] of ABB IRB 5400-22
      - target Target 220 (Cartesian target) at (1496.13, 1323.18, 1188.33) mm, rotated rx 176.39 ry 37.74 rz -142.53 deg; joints [-48.06, -13.43, 35.96, -6.9, 7.24, 5.46] of ABB IRB 5400-22
      - target Target 221 (Cartesian target) at (1572.91, 1440.71, 1166.01) mm, rotated rx 176.53 ry 36.34 rz -141.47 deg; joints [-47.09, -6.06, 30, -6.9, 7.24, 5.46] of ABB IRB 5400-22
      - target Target 222 (Cartesian target) at (1636.97, 1500.26, 1143.04) mm, rotated rx 176.61 ry 35.48 rz -141.43 deg; joints [-47.09, -1.37, 26.17, -6.9, 7.24, 5.46] of ABB IRB 5400-22
      - target Target 223 (Cartesian target) at (1811.37, 1662.37, 1168.08) mm, rotated rx 176.5 ry 36.67 rz -141.49 deg; joints [-47.09, 9.35, 14.26, -6.9, 7.24, 5.46] of ABB IRB 5400-22
      - target Target 227 (Cartesian target) at (1972.43, 1812.1, 1165.85) mm, rotated rx 176.36 ry 38.11 rz -141.57 deg; joints [-47.09, 19.39, 2.77, -6.89, 7.23, 5.45] of ABB IRB 5400-22
      - target Target 228 (Cartesian target) at (2172.53, 1998.75, 1170.16) mm, rotated rx 176 ry 41.54 rz -141.8 deg; joints [-47.08, 32.12, -13.4, -6.88, 7.23, 5.44] of ABB IRB 5400-22
      - target Target 229 (Cartesian target) at (2103.92, 2070.72, 1170.62) mm, rotated rx 176.01 ry 41.55 rz -139.86 deg; joints [-45.15, 32.11, -13.4, -6.87, 7.22, 5.43] of ABB IRB 5400-22
      - target Target 230 (Cartesian target) at (1848.91, 1880.68, 1175.31) mm, rotated rx 176.38 ry 38 rz -138.64 deg; joints [-44.17, 17.38, 4.89, -6.87, 7.22, 5.43] of ABB IRB 5400-22
      - target Target 231 (Cartesian target) at (1705.59, 1733.15, 1174.68) mm, rotated rx 176.5 ry 36.73 rz -138.57 deg; joints [-44.17, 8.01, 15.53, -6.87, 7.22, 5.43] of ABB IRB 5400-22
      - target Target 232 (Cartesian target) at (1516.46, 1538.45, 1166.57) mm, rotated rx 176.55 ry 36.28 rz -138.54 deg; joints [-44.17, -4.72, 28.72, -6.87, 7.22, 5.43] of ABB IRB 5400-22
      - target Target 233 (Cartesian target) at (1363.33, 1380.82, 1130.07) mm, rotated rx 176.54 ry 36.36 rz -138.55 deg; joints [-44.17, -15.44, 39.36, -6.87, 7.22, 5.43] of ABB IRB 5400-22
      - target Target 234 (Cartesian target) at (1163.88, 1175.5, 1127.57) mm, rotated rx 176.12 ry 40.56 rz -138.81 deg; joints [-44.17, -32.85, 52.55, -6.87, 7.22, 5.43] of ABB IRB 5400-22
      - target Target 235 (Cartesian target) at (1463.63, 1588.96, 1166.91) mm, rotated rx 176.55 ry 36.29 rz -136.61 deg; joints [-42.23, -4.72, 28.71, -6.86, 7.22, 5.42] of ABB IRB 5400-22
      - target Target 236 (Cartesian target) at (1649.3, 1793.43, 1189.09) mm, rotated rx 176.47 ry 37.15 rz -136.66 deg; joints [-42.23, 8.01, 15.11, -6.85, 7.22, 5.41] of ABB IRB 5400-22
      - target Target 237 (Cartesian target) at (1777, 1934.12, 1187.7) mm, rotated rx 176.36 ry 38.24 rz -136.73 deg; joints [-42.23, 16.71, 5.32, -6.85, 7.22, 5.41] of ABB IRB 5400-22
      - target Target 238 (Cartesian target) at (1934.66, 2107.81, 1144.83) mm, rotated rx 176.22 ry 39.61 rz -136.82 deg; joints [-42.23, 28.1, -7.45, -6.85, 7.22, 5.41] of ABB IRB 5400-22
      - target Target 239 (Cartesian target) at (2025.03, 2120.83, 1100.9) mm, rotated rx -93.18 ry 12.46 rz -115.11 deg; joints [-34.47, 42.83, -17.66, -6.84, 20.97, -86.21] of ABB IRB 5400-22
      - target Target 240 (Cartesian target) at (1760.25, 1890.55, 1106.19) mm, rotated rx -92.88 ry 14.1 rz -115.04 deg; joints [-31.59, 27.615, 5.787, -36.828, 44.685, -70.009] of ABB IRB 5400-22
      - target Target 241 (Cartesian target) at (1505.5, 1667.67, 1097.06) mm, rotated rx -92.66 ry 15.83 rz -114.98 deg; joints [-28.282, 14.511, 24.37, -49.546, 59.049, -65.394] of ABB IRB 5400-22
      - target Target 242 (Cartesian target) at (1319.72, 1459.62, 1112.1) mm, rotated rx -92.61 ry 18.73 rz -114.95 deg; joints [-25.83, 2.65, 38.07, -56.14, 68, -63.73] of ABB IRB 5400-22
      - target Target 243 (Cartesian target) at (1233.15, 1274.03, 1083.44) mm, rotated rx -92.59 ry 20.26 rz -114.94 deg; joints [-25.87, -6.06, 48.34, -60.93, 72.77, -61.87] of ABB IRB 5400-22
      - target Target 244 (Cartesian target) at (1203.49, 1210.17, 1057.53) mm, rotated rx -92.59 ry 20.27 rz -114.94 deg; joints [-25.898, -8.828, 52.011, -62.306, 74.165, -61.373] of ABB IRB 5400-22
      - target Target 245 (Cartesian target) at (1238.48, 1284.52, 1003.34) mm, rotated rx -92.66 ry 17.1 rz -114.96 deg; joints [-25.875, -3.256, 48.829, -61.115, 72.959, -61.792] of ABB IRB 5400-22
      - target Target 246 (Cartesian target) at (1246.54, 1301.68, 942.2) mm, rotated rx -92.7 ry 14.55 rz -114.97 deg; joints [-25.869, -0.52, 48.575, -61.012, 72.851, -61.826] of ABB IRB 5400-22
      - target Target 247 (Cartesian target) at (1268.69, 1349.2, 836.24) mm, rotated rx -92.78 ry 10.05 rz -114.98 deg; joints [-25.85, 5.25, 46.844, -60.299, 72.133, -62.081] of ABB IRB 5400-22
      - target Target 248 (Cartesian target) at (1288.44, 1391.28, 770.5) mm, rotated rx -92.83 ry 7.29 rz -114.99 deg; joints [-25.841, 9.431, 44.855, -59.423, 71.259, -62.403] of ABB IRB 5400-22
      - target Target 249 (Cartesian target) at (1299.86, 1415.82, 739.9) mm, rotated rx -92.85 ry 6.03 rz -114.98 deg; joints [-25.835, 11.569, 43.602, -58.85, 70.68, -62.616] of ABB IRB 5400-22
      - target Target 250 (Cartesian target) at (1429.12, 1598.7, 736.18) mm, rotated rx -92.88 ry 5.23 rz -114.98 deg; joints [-27.1, 20.06, 32.25, -53.9, 64.35, -64.22] of ABB IRB 5400-22
      - target Target 251 (Cartesian target) at (1548.08, 1736.56, 738.73) mm, rotated rx -92.91 ry 4.92 rz -114.98 deg; joints [-28.45, 26.5, 22.63, -48.83, 58.09, -66.04] of ABB IRB 5400-22
      - target Target 252 (Cartesian target) at (1728.99, 1900.56, 744.39) mm, rotated rx -92.94 ry 4.7 rz -114.97 deg; joints [-30.72, 35, 9.05, -40.02, 47.97, -69.62] of ABB IRB 5400-22
      - target Target 253 (Cartesian target) at (1779.48, 2008.97, 754.21) mm, rotated rx -92.94 ry 4.7 rz -114.97 deg; joints [-30.537, 39.366, 1.473, -32.709, 42.419, -73.619] of ABB IRB 5400-22
      - target Target 254 (Cartesian target) at (1853.63, 2073.58, 759.54) mm, rotated rx -92.94 ry 4.7 rz -114.97 deg; joints [-31.389, 43.05, -4.881, -26.342, 36.817, -76.954] of ABB IRB 5400-22
      - target Target 255 (Cartesian target) at (1933.19, 2093.91, 887.14) mm, rotated rx -92.62 ry 7.57 rz -114.92 deg; joints [-32.827, 43.02, -9.752, -20.931, 31.504, -79.534] of ABB IRB 5400-22
      - target Target 256 (Cartesian target) at (2012.01, 2090.05, 986.49) mm, rotated rx -92.32 ry 9.74 rz -114.87 deg; joints [-34.491, 43.124, -13.606, -15.874, 26.371, -81.787] of ABB IRB 5400-22
      - target Target 257 (Cartesian target) at (1973, 2075.9, 977.87) mm, rotated rx -96.03 ry 11.47 rz -123.12 deg; joints [-32.942, 44.328, -16.205, -12.339, 34.282, -84.875] of ABB IRB 5400-22
      - target Target 258 (Cartesian target) at (1952.94, 2045.31, 947.56) mm, rotated rx -96.04 ry 10.95 rz -123.12 deg; joints [-32.87, 43.132, -13.105, -16.112, 36.803, -82.436] of ABB IRB 5400-22
      - target Target 259 (Cartesian target) at (1940.23, 2026.69, 925.17) mm, rotated rx -96.05 ry 10.55 rz -123.11 deg; joints [-32.82, 42.5, -11.22, -18.29, 38.29, -81.04] of ABB IRB 5400-22
      - target Target 260 (Cartesian target) at (1888.36, 2002.28, 910.49) mm, rotated rx -96.04 ry 10.34 rz -123.1 deg; joints [-32.032, 40.603, -7.573, -22.055, 41.681, -79.021] of ABB IRB 5400-22
      - target Target 261 (Cartesian target) at (1830.88, 2022.99, 864.58) mm, rotated rx -99.01 ry 10.85 rz -125.72 deg; joints [-30.406, 41.387, -7.865, -21.188, 45.39, -78.214] of ABB IRB 5400-22
      - target Target 262 (Cartesian target) at (1786.81, 1962.77, 791.49) mm, rotated rx -98.89 ry 9.4 rz -125.7 deg; joints [-30.131, 39.799, -2.329, -26.281, 49.301, -75.024] of ABB IRB 5400-22
      - target Target 263 (Cartesian target) at (1784.33, 1958.61, 857.21) mm, rotated rx -99.05 ry 11.04 rz -125.73 deg; joints [-30.13, 38.15, -2.32, -26.28, 49.3, -75.02] of ABB IRB 5400-22
      - target Target 264 (Cartesian target) at (1781.71, 1954.08, 910.7) mm, rotated rx -99.19 ry 12.37 rz -125.76 deg; joints [-30.13, 36.81, -2.32, -26.28, 49.3, -75.02] of ABB IRB 5400-22
      - target Target 265 (Cartesian target) at (1781.71, 1954.08, 910.7) mm, rotated rx -99.19 ry 12.37 rz -125.76 deg; joints [-30.13, 36.81, -2.32, -26.28, 49.3, -75.02] of ABB IRB 5400-22
      - target Target 266 (Cartesian target) at (1861.6, 1896.03, 930.29) mm, rotated rx -99.24 ry 13.25 rz -125.76 deg; joints [-32.53, 36.14, -1.94, -27.7, 47.79, -73] of ABB IRB 5400-22
      - target Target 267 (Cartesian target) at (1699.12, 1728.06, 994.04) mm, rotated rx -70.87 ry 0.33 rz -126.34 deg; joints [-31.52, 30.5, 12.45, -44.02, 61.43, -95.19] of ABB IRB 5400-22
      - target Target 268 (Cartesian target) at (1450.31, 1445.62, 980.41) mm, rotated rx -70.87 ry 0.33 rz -126.34 deg; joints [-29.236, 16.605, 32.995, -53.385, 72.653, -91.491] of ABB IRB 5400-22
      - target Target 269 (Cartesian target) at (1405.31, 1500.09, 836.17) mm, rotated rx -70.36 ry -3.75 rz -126.34 deg; joints [-27.085, 21.872, 32.683, -53.422, 75.109, -92.056] of ABB IRB 5400-22
      - target Target 270 (Cartesian target) at (1378.56, 1464.06, 839.34) mm, rotated rx -70.36 ry -3.75 rz -126.34 deg; joints [-26.826, 20.147, 34.985, -54.114, 76.081, -91.81] of ABB IRB 5400-22
      - target Target 271 (Cartesian target) at (1376.21, 1459.8, 879.88) mm, rotated rx -70.61 ry -2.33 rz -126.32 deg; joints [-26.82, 18.72, 34.98, -54.11, 76.08, -91.8] of ABB IRB 5400-22
      - target Target 272 (Cartesian target) at (1361.34, 1439.75, 881.01) mm, rotated rx -70.61 ry -2.33 rz -126.32 deg; joints [-26.671, 17.754, 36.247, -54.463, 76.597, -91.684] of ABB IRB 5400-22
      - target Target 273 (Cartesian target) at (1356.63, 1430.46, 947.4) mm, rotated rx -71.01 ry 0.03 rz -126.31 deg; joints [-26.67, 15.37, 36.24, -54.46, 76.59, -91.68] of ABB IRB 5400-22
      - target Target 274 (Cartesian target) at (1311.33, 1441.61, 904.29) mm, rotated rx -92.76 ry 11.83 rz -114.96 deg; joints [-25.82, 7.34, 41.34, -57.77, 69.6, -63.03] of ABB IRB 5400-22
      - target Target 275 (Cartesian target) at (1326.82, 1474.47, 815.76) mm, rotated rx -92.83 ry 8.48 rz -114.97 deg; joints [-25.817, 11.553, 40.075, -57.131, 68.968, -63.268] of ABB IRB 5400-22
      - target Target 276 (Cartesian target) at (1338.35, 1499.75, 787.13) mm, rotated rx -92.85 ry 7.34 rz -114.96 deg; joints [-25.807, 13.549, 38.798, -56.48, 68.32, -63.52] of ABB IRB 5400-22
      - target Target 277 (Cartesian target) at (1315.34, 1450.29, 780.1) mm, rotated rx -92.85 ry 7.34 rz -114.96 deg; joints [-25.815, 11.653, 41.588, -57.883, 69.704, -62.963] of ABB IRB 5400-22
      - target Target 278 (Cartesian target) at (1299.2, 1416.25, 856.59) mm, rotated rx -92.81 ry 10.32 rz -114.95 deg; joints [-25.815, 7.636, 43.089, -58.603, 70.418, -62.68] of ABB IRB 5400-22
      - target Target 279 (Cartesian target) at (1295.13, 1408.32, 918.57) mm, rotated rx -92.78 ry 12.64 rz -114.93 deg; joints [-25.81, 5.33, 43.08, -58.6, 70.41, -62.67] of ABB IRB 5400-22
      - target Target 280 (Cartesian target) at (1276.13, 1368.36, 966.36) mm, rotated rx -92.75 ry 14.77 rz -114.91 deg; joints [-25.81, 1.98, 44.82, -59.4, 71.21, -62.36] of ABB IRB 5400-22
      - target Target 281 (Cartesian target) at (1260.16, 1334.08, 977.07) mm, rotated rx -92.74 ry 15.54 rz -114.91 deg; joints [-25.82, -0.03, 46.55, -60.16, 71.97, -62.07] of ABB IRB 5400-22
      - target Target 282 (Cartesian target) at (908.9, 1594.27, 977.01) mm, rotated rx -92.74 ry 15.54 rz -101.23 deg; joints [-12.14, -0.03, 46.55, -60.15, 71.96, -62.07] of ABB IRB 5400-22
      - target Target 283 (Cartesian target) at (2070.08, 2215.52, 791.95) mm, rotated rx -107.39 ry 38.45 rz -125.84 deg; joints [-32.56, 57.57, -27.53, -59.28, 74, -48.93] of ABB IRB 5400-22
      - target Target 284 (Cartesian target) at (2101.33, 2278.09, 778.09) mm, rotated rx -106.14 ry 39.47 rz -123.89 deg; joints [-32.56, 61.59, -33.4, -59.28, 72.23, -48.93] of ABB IRB 5400-22
      - target Target 285 (Cartesian target) at (2025.61, 2145.55, 808.99) mm, rotated rx -107.2 ry 35.75 rz -125.71 deg; joints [-32.57, 52.5, -20.12, -58.74, 73.43, -49.12] of ABB IRB 5400-22
      - target Target 286 (Cartesian target) at (1987.19, 2146.42, 761.12) mm, rotated rx -107.03 ry 32.97 rz -125.6 deg; joints [-31.86, 52.21, -18.25, -56.72, 72.12, -50.37] of ABB IRB 5400-22
      - target Target 287 (Cartesian target) at (2075.93, 2289.21, 711.73) mm, rotated rx -107.43 ry 37.82 rz -125.83 deg; joints [-31.86, 62.93, -33.83, -56.72, 72.12, -50.37] of ABB IRB 5400-22
      - target Target 288 (Cartesian target) at (2076, 2289.32, 615.59) mm, rotated rx -107.26 ry 35.82 rz -125.73 deg; joints [-31.86, 64.94, -33.83, -56.72, 72.12, -50.37] of ABB IRB 5400-22
      - target Target 289 (Cartesian target) at (1962.53, 2198.09, 671.07) mm, rotated rx -106.93 ry 31.77 rz -125.55 deg; joints [-30.805, 55.688, -20.66, -56.184, 72.688, -51.261] of ABB IRB 5400-22
      - target Target 290 (Cartesian target) at (1927.38, 2139.65, 701.96) mm, rotated rx -106.8 ry 30.37 rz -125.47 deg; joints [-30.8, 51.54, -15.11, -56.18, 72.68, -51.26] of ABB IRB 5400-22
      - target Target 291 (Cartesian target) at (1919.12, 2125.79, 666.73) mm, rotated rx -106.68 ry 29.09 rz -125.41 deg; joints [-30.8, 51.54, -13.83, -56.18, 72.68, -51.26] of ABB IRB 5400-22
      - target Target 292 (Cartesian target) at (1967.28, 2193.87, 682.92) mm, rotated rx -106.63 ry 28.42 rz -125.38 deg; joints [-31.01, 54.89, -20.66, -49.88, 66.37, -53.93] of ABB IRB 5400-22
      - target Target 293 (Cartesian target) at (2072.23, 2274.75, 611.72) mm, rotated rx -106.9 ry 31.41 rz -125.51 deg; joints [-32.02, 63.512, -32.209, -50.241, 65.668, -53.105] of ABB IRB 5400-22
      - target Target 294 (Cartesian target) at (1865.62, 2135.42, 645.71) mm, rotated rx -106.41 ry 24.17 rz -125.28 deg; joints [-29.72, 50.585, -12.58, -48.554, 66.568, -55.116] of ABB IRB 5400-22
      - target Target 295 (Cartesian target) at (1275.09, 1600.11, 635.02) mm, rotated rx -104.81 ry 7.06 rz -124.8 deg; joints [-21.87, 20.73, 31.3, -39.76, 67.34, -61.43] of ABB IRB 5400-22
      - target Target 296 (Cartesian target) at (1105.11, 1355.75, 598.35) mm, rotated rx -104.81 ry 7.06 rz -124.79 deg; joints [-19.148, 11.273, 46.11, -46.06, 75.976, -58.233] of ABB IRB 5400-22
      - target Target 297 (Cartesian target) at (1101.68, 1346.68, 486.89) mm, rotated rx -103.53 ry 2.47 rz -124.68 deg; joints [-19.14, 16.04, 46.11, -46.05, 75.97, -58.23] of ABB IRB 5400-22
      - target Target 298 (Cartesian target) at (1383.67, 1749.56, 516.77) mm, rotated rx -96.15 ry -1.9 rz -124.1 deg; joints [-23.048, 32.911, 20.896, -34.301, 61.497, -72.804] of ABB IRB 5400-22
      - target Target 299 (Cartesian target) at (1977.79, 2256.02, 527.36) mm, rotated rx -96.27 ry -0.64 rz -124.08 deg; joints [-31.245, 61.352, -28.914, 11.75, 23.044, -102.23] of ABB IRB 5400-22
      - target Target 300 (Cartesian target) at (2106.55, 2295.54, 516.9) mm, rotated rx -96.27 ry -0.64 rz -124.08 deg; joints [-33.575, 67.369, -38.798, 46.706, 0.953, -124.658] of ABB IRB 5400-22
      - target Target 301 (Cartesian target) at (2104.85, 2293.47, 472.08) mm, rotated rx -96.26 ry -1.57 rz -124.07 deg; joints [-33.57, 68.29, -38.79, 46.7, 0.95, -124.65] of ABB IRB 5400-22
      - target Target 302 (Cartesian target) at (1898.87, 2184.82, 478.42) mm, rotated rx -96.26 ry -1.82 rz -124.06 deg; joints [-30.35, 57.57, -20.28, -0.93, 31.1, -93.51] of ABB IRB 5400-22
      - target Target 303 (Cartesian target) at (1559.93, 1843, 461.01) mm, rotated rx -96.09 ry -2.99 rz -124.06 deg; joints [-26.523, 40.118, 11.466, -30.064, 54.398, -74.83] of ABB IRB 5400-22
      - target Target 304 (Cartesian target) at (1269.38, 1536.93, 467.76) mm, rotated rx -95.92 ry -3.77 rz -124.06 deg; joints [-22.195, 26.729, 33.576, -40.81, 67.808, -68.714] of ABB IRB 5400-22
      - target Target 305 (Cartesian target) at (1108.84, 1368.03, 446.18) mm, rotated rx -95.48 ry -5.42 rz -124.1 deg; joints [-18.92, 20.73, 44.26, -43.13, 73.42, -67.38] of ABB IRB 5400-22
      - target Target 306 (Cartesian target) at (1030.64, 1252.76, 459.44) mm, rotated rx -95.48 ry -5.41 rz -124.09 deg; joints [-17.371, 15.617, 50.89, -44.192, 76.059, -66.651] of ABB IRB 5400-22
      - target Target 307 (Cartesian target) at (1063.51, 1246.99, 743.4) mm, rotated rx -99.4 ry 7.66 rz -124.16 deg; joints [-18.737, 1.866, 51.33, -45.153, 75.431, -65.756] of ABB IRB 5400-22
      - target Target 309 (Cartesian target) at (1131.91, 1347.93, 787.14) mm, rotated rx -99.74 ry 8.78 rz -124.18 deg; joints [-20.02, 5.33, 45.37, -43.8, 72.76, -66.16] of ABB IRB 5400-22
      - target Target 309 (Cartesian target) at (1164.25, 1398.69, 696.58) mm, rotated rx -98.75 ry 4.88 rz -124.06 deg; joints [-20.519, 11.312, 42.705, -43.036, 71.521, -66.503] of ABB IRB 5400-22
      - target Target 310 (Cartesian target) at (1055.32, 1237.93, 680.24) mm, rotated rx -98.75 ry 4.88 rz -124.05 deg; joints [-18.541, 4.149, 52.02, -45.122, 75.589, -65.656] of ABB IRB 5400-22
      - target Target 311 (Cartesian target) at (645.13, 1493.57, 680.59) mm, rotated rx -98.76 ry 4.9 rz -106.97 deg; joints [-1.459, 4.14, 52.01, -45.12, 75.58, -65.65] of ABB IRB 5400-22
      - target Home (Cartesian target) at (2370, 0, 2023) mm, rotated rx 180 ry 60 rz -180 deg; joints [-90, 0, 0, -0.001, 0, 0.001] of ABB IRB 5400-22
      - target Top_Rear_Right (Cartesian target) at (2105.65, 409.3, 1463.4) mm, rotated rx -180 ry 44.94 rz -169 deg; joints [-79, -9.41, 24.47, 0, 0, 0] of ABB IRB 5400-22
      - target Target 314 (Cartesian target) at (2504.13, 901.54, 1448.4) mm, rotated rx -180 ry 45.27 rz -160.2 deg; joints [-70.2, 15.37, -0.64, 0, 0, 0] of ABB IRB 5400-22
      - target Target 315 (Cartesian target) at (2478.01, 789.4, 1508.6) mm, rotated rx -180 ry 46.49 rz -162.33 deg; joints [-72.33, 12.02, 1.49, 0, 0, 0] of ABB IRB 5400-22
      - target Target 316 (Cartesian target) at (2436.67, 731.04, 1507.87) mm, rotated rx -180 ry 46.18 rz -163.3 deg; joints [-73.3, 9.35, 4.47, 0, 0, 0] of ABB IRB 5400-22
      - target Target 317 (Cartesian target) at (2319.42, 611.09, 1488.25) mm, rotated rx -180 ry 45.22 rz -165.24 deg; joints [-75.24, 2.65, 12.13, 0, 0, 0] of ABB IRB 5400-22
      - target Target 318 (Cartesian target) at (2195.91, 345.05, 1520.33) mm, rotated rx -180 ry 46.27 rz -171.07 deg; joints [-81.07, -6.06, 19.79, 0, 0, 0] of ABB IRB 5400-22
      - target Target 320 (Cartesian target) at (2268.54, 317.21, 1512.46) mm, rotated rx -180 ry 45.9 rz -172.04 deg; joints [-82.04, -2.71, 16.81, 0, 0, 0] of ABB IRB 5400-22
      - target Target 320 (Cartesian target) at (2585.39, 728.18, 1511.83) mm, rotated rx -180 ry 47.15 rz -164.27 deg; joints [-74.27, 16.04, -3.19, 0, 0, 0] of ABB IRB 5400-22
      - target Target 321 (Cartesian target) at (2662.08, 653.38, 1505.83) mm, rotated rx -180 ry 47.45 rz -166.21 deg; joints [-76.21, 18.72, -6.17, 0, 0, 0] of ABB IRB 5400-22
      - target Roof (Cartesian target) at (2413.94, 213.32, 1469.16) mm, rotated rx -180 ry 44.73 rz -174.95 deg; joints [-84.95, 3.99, 11.28, 0, 0, 0] of ABB IRB 5400-22
      - target Target 323 (Cartesian target) at (2507.7, 136.25, 1483.89) mm, rotated rx -180 ry 45.39 rz -176.89 deg; joints [-86.89, 8.01, 6.6, 0, 0, 0] of ABB IRB 5400-22
      - target Target 324 (Cartesian target) at (2827.72, 493.52, 1563.83) mm, rotated rx -180 ry 50.36 rz -170.1 deg; joints [-80.1, 24.75, -15.11, 0, 0, 0] of ABB IRB 5400-22
      - target Target 325 (Cartesian target) at (2971.01, 313.31, 1579.13) mm, rotated rx -180 ry 52.41 rz -173.98 deg; joints [-83.98, 30.78, -23.19, 0, 0, 0] of ABB IRB 5400-22
      - target Target 326 (Cartesian target) at (2646.68, -36.03, 1533.87) mm, rotated rx -180 ry 47.46 rz 179.22 deg; joints [-90.78, 14.03, -1.49, 0, 0, 0] of ABB IRB 5400-22
      - target Target 327 (Cartesian target) at (2791.79, -227.56, 1543.38) mm, rotated rx -180 ry 49.03 rz 175.34 deg; joints [-94.66, 21.4, -10.43, 0, 0, 0] of ABB IRB 5400-22
      - target Home (Cartesian target) at (2370, 0, 2023) mm, rotated rx 180 ry 60 rz -180 deg; joints [-90, 0, 0, 0.001, -0.001, 0] of ABB IRB 5400-22
      - target Front_Side (Cartesian target) at (2904.64, 1494.98, 1065.5) mm, rotated rx 175.77 ry 45.58 rz -156.66 deg; joints [-62.62, 50.2, -35.53, -7.45, 6.69, 6.22] of ABB IRB 5400-22
      - target Target 330 (Cartesian target) at (2662.08, 1407.55, 1029.36) mm, rotated rx 176.38 ry 38.93 rz -155.59 deg; joints [-62.1, 36.9, -15.87, -0.82, 2.48, 2.26] of ABB IRB 5400-22
      - target Target 331 (Cartesian target) at (2260.19, 1139.78, 1046.74) mm, rotated rx 176.78 ry 33.57 rz -156.45 deg; joints [-63.2, 14.7, 11.7, -0.81, 2.47, 2.25] of ABB IRB 5400-22
      - target Target 332 (Cartesian target) at (2005.49, 808.42, 1033.08) mm, rotated rx 176.89 ry 32.01 rz -161.19 deg; joints [-68, -2.04, 30, -0.8, 2.46, 2.24] of ABB IRB 5400-22
      - target Target 333 (Cartesian target) at (1836.18, 383.19, 1053.03) mm, rotated rx 176.75 ry 34.23 rz -171.42 deg; joints [-78.16, -17.45, 43.19, -0.79, 2.45, 2.23] of ABB IRB 5400-22
      - target Target 335 (Cartesian target) at (1728.14, 647.06, 1064.15) mm, rotated rx 176.71 ry 34.95 rz -162.71 deg; joints [-69.42, -19.45, 44.47, -0.78, 2.44, 2.22] of ABB IRB 5400-22
      - target Target 336 (Cartesian target) at (1838.78, 688.61, 1030.22) mm, rotated rx 176.86 ry 32.7 rz -162.62 deg; joints [-69.42, -12.09, 39.36, -0.78, 2.44, 2.22] of ABB IRB 5400-22
      - target Target 336 (Cartesian target) at (2024.8, 961.31, 989.87) mm, rotated rx 177 ry 30.72 rz -157.69 deg; joints [-64.56, 2.65, 26.6, -0.77, 2.43, 2.21] of ABB IRB 5400-22
      - target Target 337 (Cartesian target) at (2144.49, 1155.18, 964.85) mm, rotated rx 177 ry 30.72 rz -154.78 deg; joints [-61.65, 12.02, 17.23, -0.77, 2.43, 2.21] of ABB IRB 5400-22
      - target Target 338 (Cartesian target) at (2641.68, 1481.65, 1002.63) mm, rotated rx 176.46 ry 38.62 rz -154.12 deg; joints [-60.68, 38.15, -16.81, -0.77, 2.43, 2.2] of ABB IRB 5400-22
      - target Target 339 (Cartesian target) at (2741.34, 1599.25, 1063.04) mm, rotated rx 176.11 ry 42.98 rz -153.37 deg; joints [-59.71, 44.84, -27.87, -0.76, 2.42, 2.19] of ABB IRB 5400-22
      - target Target 340 (Cartesian target) at (2667.03, 1679.41, 973.77) mm, rotated rx 176.33 ry 40.45 rz -151.28 deg; joints [-57.77, 44.83, -25.32, -0.75, 2.41, 2.18] of ABB IRB 5400-22
      - target Target 341 (Cartesian target) at (2197.5, 1435.94, 1017.59) mm, rotated rx 176.84 ry 33.56 rz -150 deg; joints [-56.8, 19.39, 7.02, -0.74, 2.4, 2.17] of ABB IRB 5400-22
      - target Target 342 (Cartesian target) at (1783.45, 1080.63, 1012.58) mm, rotated rx 176.98 ry 31.53 rz -151.86 deg; joints [-58.74, -5.39, 33.83, -0.73, 2.39, 2.16] of ABB IRB 5400-22
      - target Target 344 (Cartesian target) at (1579.4, 591.21, 1011.99) mm, rotated rx 176.72 ry 35.58 rz -162.68 deg; joints [-69.42, -28.16, 52.55, -0.71, 2.37, 2.14] of ABB IRB 5400-22
      - target Target 344 (Cartesian target) at (1459.29, 785.45, 985.86) mm, rotated rx 176.75 ry 35.21 rz -154.89 deg; joints [-61.65, -29.5, 54.26, -0.71, 2.37, 2.14] of ABB IRB 5400-22
      - target Target 345 (Cartesian target) at (1690.25, 1188.04, 970.39) mm, rotated rx 177.07 ry 30.25 rz -147.92 deg; joints [-54.85, -5.39, 35.11, -0.71, 2.37, 2.14] of ABB IRB 5400-22
      - target Target 346 (Cartesian target) at (2111.89, 1484.94, 986.07) mm, rotated rx 176.95 ry 32.35 rz -147.98 deg; joints [-54.85, 18.05, 9.57, -0.7, 2.36, 2.13] of ABB IRB 5400-22
      - target Target 347 (Cartesian target) at (2532.03, 1780.78, 956.3) mm, rotated rx 176.5 ry 38.85 rz -148.24 deg; joints [-54.85, 42.17, -21.06, -0.69, 2.35, 2.12] of ABB IRB 5400-22
      - target Target 348 (Cartesian target) at (2337.77, 1892.95, 897.49) mm, rotated rx 176.73 ry 35.83 rz -144.22 deg; joints [-50.97, 38.82, -14.68, -0.68, 2.34, 2.11] of ABB IRB 5400-22
      - target Target 349 (Cartesian target) at (1914.74, 1604.48, 936.09) mm, rotated rx 177.1 ry 30.35 rz -143.04 deg; joints [-50, 15.36, 14.26, -0.66, 2.32, 2.09] of ABB IRB 5400-22
      - target Target 350 (Cartesian target) at (1586.43, 1328.96, 949.71) mm, rotated rx 177.12 ry 29.59 rz -143.04 deg; joints [-50, -4.72, 35.11, -0.7, 2.36, 2.13] of ABB IRB 5400-22
      - target Target 351 (Cartesian target) at (1395.35, 946.6, 945.07) mm, rotated rx 176.76 ry 35.21 rz -149.07 deg; joints [-54.779, -26.644, 54.41, -26.664, 19.942, 17.017] of ABB IRB 5400-22
      - target Target 352 (Cartesian target) at (1322.76, 1066.74, 874.65) mm, rotated rx 176.76 ry 35.2 rz -144.43 deg; joints [-49.519, -23.862, 55.874, -41.968, 31.708, 24.82] of ABB IRB 5400-22
      - target Target 353 (Cartesian target) at (1571.28, 1494.48, 869.88) mm, rotated rx 176.78 ry 35.21 rz -139.43 deg; joints [-45.15, 1.81, 35.14, -55.63, 42.35, 31.26] of ABB IRB 5400-22
      - target Target 354 (Cartesian target) at (1947.54, 1804.91, 896.42) mm, rotated rx 176.47 ry 38.5 rz -140.58 deg; joints [-46.147, 22.789, 10.286, -54.346, 41.169, 30.762] of ABB IRB 5400-22
      - target Target 355 (Cartesian target) at (2221.34, 1995.49, 848.2) mm, rotated rx 176.78 ry 35.15 rz -141.27 deg; joints [-47.728, 38.583, -12.496, -17.064, 12.854, 11.827] of ABB IRB 5400-22
      - target Target 356 (Cartesian target) at (2133.25, 2030.51, 819.37) mm, rotated rx 176.79 ry 35.14 rz -139.66 deg; joints [-45.854, 37.147, -8.976, -28.894, 20.958, 18.497] of ABB IRB 5400-22
      - target Target 357 (Cartesian target) at (1975.23, 1909.46, 857.65) mm, rotated rx 176.79 ry 35.16 rz -139.29 deg; joints [-45.15, 27.56, 3.7, -40.42, 29.65, 24.45] of ABB IRB 5400-22
      - target Target 358 (Cartesian target) at (1801, 1848.92, 850.77) mm, rotated rx 176.79 ry 35.16 rz -137.66 deg; joints [-43.2, 20.52, 13.78, -48.85, 36.73, 28.28] of ABB IRB 5400-22
      - target Target 359 (Cartesian target) at (1521.05, 1589.55, 845.12) mm, rotated rx 176.8 ry 35.17 rz -137.43 deg; joints [-42.23, 3.94, 34.02, -56.66, 44.39, 31.13] of ABB IRB 5400-22
      - target Target 360 (Cartesian target) at (1368.57, 1412.18, 820.82) mm, rotated rx 176.8 ry 35.16 rz -138.04 deg; joints [-42.23, -6.69, 45.53, -57.82, 46.19, 31.23] of ABB IRB 5400-22
      - target Target 361 (Cartesian target) at (1295.42, 1147.05, 843.49) mm, rotated rx 176.81 ry 35.16 rz -142.67 deg; joints [-46.367, -20.881, 55.34, -47.051, 37.378, 26.453] of ABB IRB 5400-22
      - target Target 362 (Cartesian target) at (1230.24, 1350.84, 744.36) mm, rotated rx 176.59 ry 36.62 rz -136.71 deg; joints [-39.97, -11.42, 53.93, -66.82, 55.9, 33.77] of ABB IRB 5400-22
      - target Target 363 (Cartesian target) at (1219.19, 1338.19, 666.59) mm, rotated rx 177.16 ry 32.63 rz -136.39 deg; joints [-40.003, -9.675, 54.333, -63.428, 52.464, 32.754] of ABB IRB 5400-22
      - target Target 364 (Cartesian target) at (1248.62, 1414.66, 685.93) mm, rotated rx 177.15 ry 32.62 rz -135.36 deg; joints [-39.29, -6.327, 50.506, -62.863, 51.523, 32.733] of ABB IRB 5400-22
      - target Target 365 (Cartesian target) at (1203.67, 1370.27, 645.5) mm, rotated rx 177.15 ry 32.62 rz -135.36 deg; joints [-38.949, -8.046, 54.047, -65.863, 54.92, 33.492] of ABB IRB 5400-22
      - target Target 366 (Cartesian target) at (1199.85, 1357.53, 595.96) mm, rotated rx -105.77 ry -15.09 rz -67.77 deg; joints [-41.165, -4.56, 56.012, -9.242, -32.694, -75.184] of ABB IRB 5400-22
      - target Target 367 (Cartesian target) at (1261.03, 1565.56, 520.66) mm, rotated rx -105.49 ry -14.92 rz -67.84 deg; joints [-36.1, 8.01, 49.11, -98.63, 35.79, -28.76] of ABB IRB 5400-22
      - target Target 368 (Cartesian target) at (1149.7, 1285.64, 589.19) mm, rotated rx -107.33 ry -15.8 rz -67.34 deg; joints [-39.83, -10.08, 62.04, -101.61, 29.63, -21.91] of ABB IRB 5400-22
      - target Target 369 (Cartesian target) at (1150.6, 1287.16, 655.77) mm, rotated rx -104.88 ry -14.55 rz -67.97 deg; joints [-39.82, -12.76, 62.04, -101.6, 29.62, -21.91] of ABB IRB 5400-22
      - target Target 370 (Cartesian target) at (1150.06, 1195.02, 593.82) mm, rotated rx -108.59 ry -16.18 rz -66.98 deg; joints [-42.97, -14.77, 64.95, -109.16, 30.47, -15.85] of ABB IRB 5400-22
      - target Target 371 (Cartesian target) at (1188.53, 1066.74, 613.34) mm, rotated rx -109.66 ry -16.49 rz -66.68 deg; joints [-49.64, -20.12, 67.56, -127.37, 36.84, -4.86] of ABB IRB 5400-22
      - target Target 372 (Cartesian target) at (1182.75, 1061.72, 508.29) mm, rotated rx -114.34 ry -17.79 rz -65.31 deg; joints [-49.64, -15.44, 67.54, -127.35, 36.84, -4.86] of ABB IRB 5400-22
      - target Target 373 (Cartesian target) at (1140.64, 1171.81, 545.28) mm, rotated rx -111.27 ry -16.6 rz -66.21 deg; joints [-43.63, -14.1, 65.82, -111.92, 31.43, -13.36] of ABB IRB 5400-22
      - target Target 374 (Cartesian target) at (1166.09, 1390.95, 542.79) mm, rotated rx -108.01 ry -14.88 rz -67.09 deg; joints [-37.57, -2.71, 58.01, -100.68, 33.32, -23.96] of ABB IRB 5400-22
      - target Target 375 (Cartesian target) at (1176.45, 1298.73, 481.02) mm, rotated rx -111.36 ry -16.44 rz -66.19 deg; joints [-40.708, -3.617, 60.598, -107.057, 34.186, -19.682] of ABB IRB 5400-22
      - target Target 376 (Cartesian target) at (1176.83, 1260.16, 381.83) mm, rotated rx -115.47 ry -18.24 rz -64.95 deg; joints [-41.953, -0.395, 61.157, -109.646, 34.747, -18.246] of ABB IRB 5400-22
      - target Target 377 (Cartesian target) at (1156.57, 1216.32, 327.88) mm, rotated rx -118.44 ry -19.4 rz -63.99 deg; joints [-42.657, -0.064, 62.573, -110.596, 33.893, -16.836] of ABB IRB 5400-22
      - target Target 378 (Cartesian target) at (1163.11, 1303.95, 346.95) mm, rotated rx -116.08 ry -18.42 rz -64.76 deg; joints [-40.1, 2.65, 59.83, -106.29, 34.54, -20.35] of ABB IRB 5400-22
      - target Target 379 (Cartesian target) at (1176.48, 1319.83, 466.28) mm, rotated rx -111.64 ry -16.41 rz -66.09 deg; joints [-40.1, -2.04, 59.83, -106.29, 34.54, -20.35] of ABB IRB 5400-22
      - target Target 380 (Cartesian target) at (1159.48, 1366.95, 482.56) mm, rotated rx -110.57 ry -15.86 rz -66.38 deg; joints [-38.09, -1.37, 58.77, -102.15, 33.62, -22.66] of ABB IRB 5400-22
      - target Target 381 (Cartesian target) at (1149.54, 1354.27, 378.46) mm, rotated rx -114.29 ry -17.74 rz -65.31 deg; joints [-38.09, 2.65, 58.77, -102.15, 33.62, -22.66] of ABB IRB 5400-22
      - target Target 382 (Cartesian target) at (1192.85, 1401.91, 342.34) mm, rotated rx -114.29 ry -17.74 rz -65.31 deg; joints [-38.309, 7.492, 55.738, -104.117, 36.295, -23.24] of ABB IRB 5400-22
      - target Target 383 (Cartesian target) at (1189.21, 1410.79, 438.83) mm, rotated rx -111.16 ry -16.17 rz -66.21 deg; joints [-37.94, 3.32, 56.25, -103.1, 35.6, -23.42] of ABB IRB 5400-22
      - target Target 384 (Cartesian target) at (1181.46, 1428.37, 433.26) mm, rotated rx -111.16 ry -16.17 rz -66.21 deg; joints [-37.193, 4.02, 55.799, -101.656, 35.302, -24.193] of ABB IRB 5400-22
      - target Target 385 (Cartesian target) at (1162.93, 1417.49, 385.56) mm, rotated rx -112.97 ry -17.12 rz -65.7 deg; joints [-36.827, 5.201, 56.31, -100.606, 34.604, -24.404] of ABB IRB 5400-22
      - target Target 386 (Cartesian target) at (1349.82, 1675.94, 371.95) mm, rotated rx -111.49 ry -16.32 rz -66.78 deg; joints [-36.41, 18.62, 41, -97.91, 33.28, -25.34] of ABB IRB 5400-22
      - target Target 387 (Cartesian target) at (1588.81, 1944.57, 389.25) mm, rotated rx -104.51 ry -3.95 rz -84 deg; joints [-33.5, 34.13, 22.34, -81.55, 44.27, -34.95] of ABB IRB 5400-22
      - target Target 388 (Cartesian target) at (1638.71, 1991.08, 389.32) mm, rotated rx -104.36 ry 9.44 rz -97.59 deg; joints [-30.91, 40.16, 15.96, -79.18, 63.66, -36.66] of ABB IRB 5400-22
      - target Target 389 (Cartesian target) at (1696.36, 2056.23, 381.1) mm, rotated rx -105.11 ry 16.92 rz -104.07 deg; joints [-30.07, 45.51, 8.72, -78.47, 72.48, -37.18] of ABB IRB 5400-22
      - target Target 390 (Cartesian target) at (1698.21, 2051.66, 485.25) mm, rotated rx -104.33 ry 19.5 rz -103.81 deg; joints [-30.171, 42.527, 9.543, -79.347, 73.349, -36.991] of ABB IRB 5400-22
      - target Target 391 (Cartesian target) at (1700.29, 2055.32, 554.28) mm, rotated rx -103.82 ry 21.12 rz -103.64 deg; joints [-30.17, 40.83, 9.54, -79.34, 73.34, -36.99] of ABB IRB 5400-22
      - target Target 392 (Cartesian target) at (1757.46, 2023.2, 530.82) mm, rotated rx -103.82 ry 21.12 rz -103.64 deg; joints [-31.881, 41.692, 9.352, -81.961, 74.237, -35.684] of ABB IRB 5400-22
      - target Target 393 (Cartesian target) at (1812.24, 2085.5, 544.68) mm, rotated rx -103.86 ry 21.03 rz -103.64 deg; joints [-32.24, 44.17, 4.19, -78.12, 69.36, -35.96] of ABB IRB 5400-22
      - target Target 394 (Cartesian target) at (1811.4, 2084.31, 516.19) mm, rotated rx -104.09 ry 20.39 rz -103.71 deg; joints [-32.24, 44.84, 4.19, -78.12, 69.35, -35.95] of ABB IRB 5400-22
      - target Target 395 (Cartesian target) at (1824.4, 2152.53, 399.56) mm, rotated rx -105.22 ry 17.21 rz -104.07 deg; joints [-31.644, 50.087, -0.757, -72.727, 64.111, -37.251] of ABB IRB 5400-22
      - target Target 396 (Cartesian target) at (1990.21, 2201.06, 393.24) mm, rotated rx -109.63 ry 30.7 rz -124.13 deg; joints [-31.55, 62.26, -21.06, -62.91, 76.89, -44.27] of ABB IRB 5400-22
      - target Target 397 (Cartesian target) at (2054.34, 2144.93, 352.21) mm, rotated rx -109.63 ry 30.7 rz -124.13 deg; joints [-33.39, 62.983, -20.423, -65.751, 77.895, -42.282] of ABB IRB 5400-22
      - target Target 398 (Cartesian target) at (2022.01, 2095.99, 454.63) mm, rotated rx -109.63 ry 29.96 rz -124.13 deg; joints [-33.399, 57.224, -14.805, -64.463, 76.51, -42.674] of ABB IRB 5400-22
      - target Target 399 (Cartesian target) at (1944.53, 2144.87, 445.04) mm, rotated rx -109.63 ry 29.96 rz -122.3 deg; joints [-31.55, 56.77, -13.49, -65.71, 77.86, -42.29] of ABB IRB 5400-22
      - target Target 400 (Cartesian target) at (1734.41, 2013.34, 532.32) mm, rotated rx -103.88 ry 21.2 rz -103.63 deg; joints [-31.506, 40.911, 10.638, -82.438, 75.252, -35.775] of ABB IRB 5400-22
      - target Target 401 (Cartesian target) at (2105.51, 2203, 594.75) mm, rotated rx -103.52 ry 22 rz -103.49 deg; joints [-36.49, 53.55, -14.47, -69.05, 54.22, -35.16] of ABB IRB 5400-22
      - target Target 402 (Cartesian target) at (2206.92, 2216.9, 595.27) mm, rotated rx -107.37 ry 34.66 rz -114.16 deg; joints [-36.49, 60.92, -25.74, -69.05, 67.57, -35.15] of ABB IRB 5400-22
      - target Target 403 (Cartesian target) at (1924.29, 2136.69, 603.82) mm, rotated rx -103.43 ry 22.22 rz -103.45 deg; joints [-33.891, 46.684, -2.656, -74.987, 63.765, -35.456] of ABB IRB 5400-22
      - target Target 404 (Cartesian target) at (1959.8, 2095.37, 660.22) mm, rotated rx -102.74 ry 23.94 rz -103.17 deg; joints [-35.153, 44.996, -1.642, -78.112, 65.677, -34.07] of ABB IRB 5400-22
      - target Target 405 (Cartesian target) at (1888.09, 2068.51, 619.05) mm, rotated rx -103.09 ry 23.12 rz -103.31 deg; joints [-34.07, 43.5, 2.58, -79.86, 69.01, -34.53] of ABB IRB 5400-22
      - target Target 406 (Cartesian target) at (1940.45, 2056.81, 692.44) mm, rotated rx -102.31 ry 24.98 rz -102.99 deg; joints [-35.303, 42.679, 1.249, -80.857, 68.614, -33.559] of ABB IRB 5400-22
      - target Target 407 (Cartesian target) at (2003.32, 2112.05, 712.35) mm, rotated rx -102.31 ry 24.98 rz -102.99 deg; joints [-35.78, 45.416, -4.391, -76.845, 63.476, -33.81] of ABB IRB 5400-22
      - target Target 408 (Cartesian target) at (2002.27, 2110.65, 768.46) mm, rotated rx -101.77 ry 26.13 rz -102.75 deg; joints [-35.78, 44.17, -4.39, -76.84, 63.47, -33.81] of ABB IRB 5400-22
      - target Target 409 (Cartesian target) at (1986.42, 2040.59, 733.23) mm, rotated rx -101.77 ry 26.13 rz -102.75 deg; joints [-36.452, 42.431, 0.265, -82.047, 68.553, -32.609] of ABB IRB 5400-22
      - target Target 411 (Cartesian target) at (1973.4, 2066.55, 719.14) mm, rotated rx -112.97 ry 31.21 rz -107.7 deg; joints [-35.901, 41.764, -0.699, -76.315, 66.835, -24.502] of ABB IRB 5400-22
      - target Target 411 (Cartesian target) at (2051.35, 2019.39, 802.5) mm, rotated rx -132.56 ry 44.47 rz -122.74 deg; joints [-37.773, 39.991, -2.734, -73.49, 73.597, -11.362] of ABB IRB 5400-22
      - target Target 412 (Cartesian target) at (2087.44, 2032.18, 826.26) mm, rotated rx -132.41 ry 45.63 rz -122.23 deg; joints [-38.35, 40.92, -4.81, -74.18, 73.27, -10.5] of ABB IRB 5400-22
      - target Target 413 (Cartesian target) at (1817.19, 1942.27, 860.06) mm, rotated rx -134.17 ry 39.64 rz -123.3 deg; joints [-34.333, 29.223, 8.868, -64.559, 67.724, -14.825] of ABB IRB 5400-22
      - target Target 414 (Cartesian target) at (1532.76, 1687.05, 867.38) mm, rotated rx -123.12 ry 29.51 rz -122.85 deg; joints [-29.77, 16.04, 25.84, -55.38, 66.75, -32.25] of ABB IRB 5400-22
      - target Target 415 (Cartesian target) at (1416.27, 1484.04, 838.65) mm, rotated rx -122.98 ry 27.07 rz -122.78 deg; joints [-29.76, 6.67, 37.66, -55.37, 66.75, -32.25] of ABB IRB 5400-22
      - target Target 416 (Cartesian target) at (1302.02, 1284.22, 834.58) mm, rotated rx -122.96 ry 26.73 rz -122.77 deg; joints [-29.76, -4.05, 48.72, -55.37, 66.75, -32.25] of ABB IRB 5400-22
      - target Target 417 (Cartesian target) at (1262.15, 1214.49, 830.83) mm, rotated rx -122.98 ry 26.92 rz -122.78 deg; joints [-29.76, -8.07, 52.55, -55.37, 66.75, -32.25] of ABB IRB 5400-22
      - target Target 418 (Cartesian target) at (1287.91, 1061.82, 853.23) mm, rotated rx -123.44 ry 31.68 rz -123.01 deg; joints [-34.33, -14.77, 58.48, -64.17, 70.55, -26.48] of ABB IRB 5400-22
      - target Target 419 (Cartesian target) at (638.08, 1542.41, 853.13) mm, rotated rx -123.46 ry 31.68 rz -94.99 deg; joints [-6.31, -14.77, 58.48, -64.16, 70.54, -26.47] of ABB IRB 5400-22
      - target Home (Cartesian target) at (2370, 0, 2023) mm, rotated rx -180 ry 60 rz -180 deg; joints [-90, 0, 0, 0.001, -0.001, 0] of ABB IRB 5400-22
      - target Top_Front_Left (Cartesian target) at (2739.69, 335.91, 1448.51) mm, rotated rx -180 ry 46.11 rz -173.01 deg; joints [-83.01, 20.06, -6.17, 0, 0, 0] of ABB IRB 5400-22
      - target Target 422 (Cartesian target) at (3279.47, 402.09, 1533.29) mm, rotated rx -180 ry 58.7 rz -173.01 deg; joints [-83.01, 50.87, -49.57, 0, 0, 0] of ABB IRB 5400-22
      - target Target 431 (Cartesian target) at (3285.31, 234.34, 1567.64) mm, rotated rx -180 ry 59.35 rz -175.92 deg; joints [-85.92, 50.2, -49.55, 0, 0, 0] of ABB IRB 5400-22
      - target Target 424 (Cartesian target) at (2757.96, 197.21, 1478.94) mm, rotated rx -180 ry 46.96 rz -175.91 deg; joints [-85.91, 20.06, -7.02, 0, 0, 0] of ABB IRB 5400-22
      - target Target 425 (Cartesian target) at (2744.61, 56.05, 1536.36) mm, rotated rx -180 ry 48.3 rz -178.83 deg; joints [-88.83, 18.72, -7.02, 0, 0, 0] of ABB IRB 5400-22
      - target Target 432 (Cartesian target) at (3270.73, 125.25, 1591.32) mm, rotated rx -177.19 ry 59.32 rz -171.03 deg; joints [-88.81, 48.86, -48.3, 2.33, -6.99, 2.33] of ABB IRB 5400-22
      - target Target 433 (Cartesian target) at (3277.85, -155.15, 1618.47) mm, rotated rx -180 ry 60.46 rz 177.29 deg; joints [-92.71, 49.53, -49.99, 0, 0, 0] of ABB IRB 5400-22
      - target Target 428 (Cartesian target) at (2756.14, -130.94, 1538.25) mm, rotated rx -180 ry 48.48 rz 177.28 deg; joints [-92.72, 19.39, -7.87, 0, 0, 0] of ABB IRB 5400-22
      - target Target 429 (Cartesian target) at (2770.39, -320.55, 1556.71) mm, rotated rx -180 ry 49.26 rz 173.4 deg; joints [-96.6, 20.73, -9.99, 0, 0, 0] of ABB IRB 5400-22
      - target Target 434 (Cartesian target) at (3225.77, -373.23, 1618.75) mm, rotated rx -180 ry 59.31 rz 173.4 deg; joints [-96.6, 46.85, -46.16, 0, 0, 0] of ABB IRB 5400-22
      - target Target 431 (Cartesian target) at (3278.35, -549.2, 1630.76) mm, rotated rx -180 ry 62.56 rz 170.49 deg; joints [-99.51, 53.4, -55.96, 0, 0, 0] of ABB IRB 5400-22
      - target Target 432 (Cartesian target) at (2789.61, -467.32, 1545.8) mm, rotated rx -180 ry 49.39 rz 170.49 deg; joints [-99.51, 22.74, -12.13, 0, 0, 0] of ABB IRB 5400-22
      - target Target 433 (Cartesian target) at (2813.32, -620.09, 1533.71) mm, rotated rx -180 ry 49.69 rz 167.57 deg; joints [-102.43, 25.42, -15.11, 0, 0, 0] of ABB IRB 5400-22
      - target Home (Cartesian target) at (2370, 0, 2023) mm, rotated rx -180 ry 60 rz -180 deg; joints [-90, 0, 0, 0.001, -0.001, 0] of ABB IRB 5400-22
      - target After-45_Top_Rear_Left (Cartesian target) at (2092.96, -424.3, 1484.92) mm, rotated rx -180 ry 45.61 rz 168.54 deg; joints [-101.46, -10.08, 24.47, 0, 0, 0] of ABB IRB 5400-22
      - target Target 436 (Cartesian target) at (2426.62, -811.93, 1511.95) mm, rotated rx -180 ry 46.36 rz 161.5 deg; joints [-108.5, 10.02, 3.62, 0, 0, 0] of ABB IRB 5400-22
      - target Target 437 (Cartesian target) at (2512.41, -735.16, 1527.45) mm, rotated rx -180 ry 47.1 rz 163.69 deg; joints [-106.31, 12.69, 0.21, 0, 0, 0] of ABB IRB 5400-22
      - target Target 438 (Cartesian target) at (2163.76, -363.13, 1498.73) mm, rotated rx -180 ry 47.13 rz 170.5 deg; joints [-98.86, -7.4, 22.34, -24.72, 16.16, 14.32] of ABB IRB 5400-22
      - target Target 439 (Cartesian target) at (2299.8, -279.42, 1490.46) mm, rotated rx 179.98 ry 46.63 rz 173.11 deg; joints [-97.57, -1.37, 16.81, 24.63, -16.15, -14.23] of ABB IRB 5400-22
      - target Target 440 (Cartesian target) at (2695.93, -642.26, 1524.89) mm, rotated rx -180 ry 48.24 rz 166.6 deg; joints [-103.4, 20.06, -8.3, 0, 0, 0] of ABB IRB 5400-22
      - target Target 441 (Cartesian target) at (2814.74, -471.53, 1532.13) mm, rotated rx -180 ry 49.32 rz 170.49 deg; joints [-99.51, 24.08, -13.4, 0, 0, 0] of ABB IRB 5400-22
      - target Target 442 (Cartesian target) at (2371.47, -167.29, 1516.55) mm, rotated rx -180 ry 47.35 rz 176.03 deg; joints [-94.66, 1.31, 13.4, 24.62, -16.14, -14.23] of ABB IRB 5400-22
      - target Target 443 (Cartesian target) at (2547.09, -51.88, 1517.72) mm, rotated rx -180 ry 47.82 rz 178.94 deg; joints [-91.75, 9.35, 4.89, 24.61, -16.13, -14.22] of ABB IRB 5400-22
      - target Target 444 (Cartesian target) at (2940.77, -340.26, 1549.45) mm, rotated rx -180 ry 51.2 rz 173.4 deg; joints [-96.6, 29.44, -20.64, 0, 0, 0] of ABB IRB 5400-22
      - target Target 445 (Cartesian target) at (3049.89, -248.6, 1573) mm, rotated rx -180 ry 53.5 rz 175.34 deg; joints [-94.66, 34.8, -28.3, 0, 0, 0] of ABB IRB 5400-22
      - target Target 446 (Cartesian target) at (2702.3, 172.79, 1554.79) mm, rotated rx -179.97 ry 49.82 rz -176.18 deg; joints [-86.89, 16.71, -4.47, 24.6, -16.12, -14.21] of ABB IRB 5400-22
      - target Home (Cartesian target) at (2370, 0, 2023) mm, rotated rx -180 ry 60 rz -180 deg; joints [-90, 0, 0, -0.001, 0.001, 0.001] of ABB IRB 5400-22
      - target Top_Front_Right (Cartesian target) at (2716.47, -296.79, 1465.16) mm, rotated rx 179.93 ry 49.54 rz 173.63 deg; joints [-96.964, 18.414, -3.006, 38.173, -25.506, -21.631] of ABB IRB 5400-22
      - target Target 449 (Cartesian target) at (3257.39, -376.89, 1514.43) mm, rotated rx -180 ry 57.29 rz 173.4 deg; joints [-96.6, 48.86, -46.15, 0, 0, 0] of ABB IRB 5400-22
      - target Target 450 (Cartesian target) at (3288.87, -155.67, 1583.18) mm, rotated rx -180 ry 59.78 rz 177.29 deg; joints [-92.71, 50.2, -49.98, 0, 0, 0] of ABB IRB 5400-22
      - target Target 451 (Cartesian target) at (2775.95, -131.4, 1480.14) mm, rotated rx -180 ry 47.13 rz 177.29 deg; joints [-92.71, 20.73, -7.86, 0, 0, 0] of ABB IRB 5400-22
      - target Target 452 (Cartesian target) at (2744.61, 56.05, 1536.36) mm, rotated rx 180 ry 48.3 rz -178.83 deg; joints [-88.83, 18.72, -7.02, 0, 0, 0] of ABB IRB 5400-22
      - target Target 453 (Cartesian target) at (3270.73, 125.25, 1591.32) mm, rotated rx -177.19 ry 59.32 rz -171.03 deg; joints [-88.81, 48.86, -48.3, 2.33, -6.99, 2.33] of ABB IRB 5400-22
      - target Target 454 (Cartesian target) at (2727.77, 195.53, 1564.89) mm, rotated rx -180 ry 48.97 rz -175.9 deg; joints [-85.9, 18.05, -7.02, 0, 0, 0] of ABB IRB 5400-22
      - target Target 455 (Cartesian target) at (3274.55, 233.57, 1602.22) mm, rotated rx -180 ry 60.01 rz -175.92 deg; joints [-85.92, 49.53, -49.54, 0, 0, 0] of ABB IRB 5400-22
      - target Target 456 (Cartesian target) at (3233.85, 564.4, 1602.38) mm, rotated rx -180 ry 60.01 rz -170.1 deg; joints [-80.1, 49.52, -49.53, 0, 0, 0] of ABB IRB 5400-22
      - target Target 457 (Cartesian target) at (2777.73, 533.4, 1545.8) mm, rotated rx -180 ry 49.39 rz -169.13 deg; joints [-79.13, 22.74, -12.13, 0, 0, 0] of ABB IRB 5400-22
      - target Home (Cartesian target) at (2370, 0, 2023) mm, rotated rx 180 ry 60 rz -180 deg; joints [-90, 0, 0, -0.001, 0.001, 0.001] of ABB IRB 5400-22
  - Python program Inspect_Car_Painting_Station (listed below)
  - Python program Prog4 (listed below)
  - Python program Car_Rotation_180 (listed below)
  - Python program Car_Rotation_90 (listed below)
  - Python program Car_Rotation_45 (listed below)
  - frame Frame 6 at (0, 2000, 0) mm
  - frame Components at (0, 0, 0) mm
    - frame Truntable 1 Frame at (3300, 0, 0) mm
      - object Turntable 1 at (0, 0, 0) mm
        - item type 7 Turntable 1-0
        - item type 7 Turntable 1-1
        - item type 7 Turntable 1-2
        - item type 7 Turntable 1-3
        - item type 7 Turntable 1-4
  - frame Car Rotary Fixture Base at (3300, 1000, 0) mm
    - robot Car Rotary Fixture: 1 axes
        modified DH rows (alpha deg, a mm, theta deg, d mm): 0, 0, 0, 0
        joint limits [0] to [360]; home [0]; saved at [180]
  - Python program Car_Rotation_-45 (listed below)
  - Python program Car_Rotation_0 (listed below)
  - Python program Full_Painting (listed below)

--- Python program Inspect_Car_Painting_Station ---
from robodk.robolink import *

RDK = Robolink()

robot = RDK.Item("ABB IRB 5400-22", ITEM_TYPE_ROBOT)
target_196 = RDK.Item("Target 196", ITEM_TYPE_TARGET)
target_197 = RDK.Item("Target 197", ITEM_TYPE_TARGET)

if not robot.Valid():
    raise Exception("Robot not found")

if not target_196.Valid() or not target_197.Valid():
    raise Exception("Target 196 or Target 197 not found")

print("Moving to Target 196...")
robot.MoveJ(target_196)

print("Testing linear movement to Target 197...")
robot.MoveL(target_197)

print("Linear movement to Target 197 succeeded.")

--- Python program Prog4 ---
# ============================================================
# YUKTII ROBOTIC CAR PAINTING CELL
# ABB IRB 5400-22
#
# COMPLETE PAINTING + ROTATION + BOUNDARY SEQUENCE
#
# PHASE 1: Initial Home
#
# PHASE 2: Original-side painting
#   Paint_Side_P01 ... Paint_Side_P59
#   Target 64 ... Target 91
#   Target 93, Target 93, Target 94
#   Target 96, Target 96, Target 97
#   Target 99, Target 99
#   Target 100 ... Target 106
#
# PHASE 3: Return to Home after Target 106
#
# PHASE 4: Slowly rotate the car by 180 degrees
#
# PHASE 5: New-side outline
#   New_Side1
#   Target 108 ... Target 138
#   Target 174, Target 175
#   Target 140 ... Target 172
#
# PHASE 6: Return to Home after Target 172
#
# PHASE 7: Additional boundary
#   Target 175 ... Target 205
#   Target 207, Target 207
#   Target 208 ... Target 212
#
# PHASE 8: Return to final Home
#
# IMPORTANT:
# - Executes movements directly in RoboDK.
# - Does not create a saved RoboDK program.
# - Validates targets before robot movement.
# ============================================================

from robodk.robolink import *
import time

RDK = Robolink()

# ------------------------------------------------------------
# CONFIGURATION
# ------------------------------------------------------------

ROBOT_NAME = "ABB IRB 5400-22"
FRAME_NAME = "Painting Cell Frame"
TOOL_NAME = "Generic Paint Sprayer"
FIXTURE_NAME = "Car Rotary Fixture"

ROTATION_DEGREES = 180.0
ROBOT_SPEED = 50

# Rotation speed: reduce STEP_ANGLE or increase STEP_DELAY
# for slower visible rotation.
STEP_ANGLE = 2.0
STEP_DELAY = 0.10

# ------------------------------------------------------------
# PHASE 0: FIND STATION ITEMS
# ------------------------------------------------------------

robot = RDK.Item(ROBOT_NAME, ITEM_TYPE_ROBOT)
frame = RDK.Item(FRAME_NAME, ITEM_TYPE_FRAME)
tool = RDK.Item(TOOL_NAME)
fixture = RDK.Item(FIXTURE_NAME)

for item, name in [
    (robot, ROBOT_NAME),
    (frame, FRAME_NAME),
    (tool, TOOL_NAME),
    (fixture, FIXTURE_NAME),
]:
    if not item.Valid():
        raise Exception("Station item not found: " + name)

# ------------------------------------------------------------
# BUILD ORIGINAL-SIDE SEQUENCE
# ------------------------------------------------------------

original_names = []

# Paint_Side_P01 through Paint_Side_P59
for i in range(1, 60):
    original_names.append(
        "Paint_Side_P" + str(i).zfill(2)
    )

# Target 64 through Target 91
for i in range(64, 92):
    original_names.append("Target " + str(i))

# Preserve duplicate occurrences in the supplied sequence.
original_names.extend([
    "Target 93",
    "Target 93",
    "Target 94",
    "Target 96",
    "Target 96",
    "Target 97",
    "Target 99",
    "Target 99",
])

# Target 100 through Target 106
for i in range(100, 107):
    original_names.append("Target " + str(i))

# ------------------------------------------------------------
# BUILD NEW-SIDE OUTLINE SEQUENCE
# ------------------------------------------------------------

outline_names = ["New_Side1"]

# Target 108 through Target 138
for i in range(108, 139):
    outline_names.append("Target " + str(i))

# These appear between Target 138 and Target 140.
outline_names.extend([
    "Target 174",
    "Target 175",
])

# Continue from Target 140 through Target 172.
for i in range(140, 173):
    outline_names.append("Target " + str(i))

# ------------------------------------------------------------
# BUILD ADDITIONAL BOUNDARY SEQUENCE
# ------------------------------------------------------------

boundary_names = []

# Target 175 through Target 205
for i in range(175, 206):
    boundary_names.append("Target " + str(i))

# Preserve the duplicate Target 207.
boundary_names.extend([
    "Target 207",
    "Target 207",
])

# Target 208 through Target 212
for i in range(208, 213):
    boundary_names.append("Target " + str(i))

# ------------------------------------------------------------
# COLLECT TARGETS AND PRESERVE OCCURRENCE ORDER
# ------------------------------------------------------------

all_targets = RDK.ItemList(ITEM_TYPE_TARGET)

targets_by_name = {}

for item in all_targets:
    if item.Valid():
        targets_by_name.setdefault(
            item.Name(), []
        ).append(item)

# The screenshots show five Home targets in tree order:
# Home 1: initial Home
# Home 2: after Paint_Side_P59
# Home 3: after Target 106
# Home 4: after Target 172
# Home 5: after Target 212

homes = targets_by_name.get("Home", [])

if len(homes) < 5:
    raise Exception(
        "Expected at least 5 Home targets in station-tree order. "
        "Found " + str(len(homes))
        + ". No robot movement has started."
    )

initial_home = homes[0]
home_after_106 = homes[2]
home_after_172 = homes[3]
final_home = homes[4]

# ------------------------------------------------------------
# RESOLVE ALL TARGETS USING SHARED DUPLICATE-NAME COUNTERS
# ------------------------------------------------------------

# Shared counters are important because Target 175 appears
# once in the outline sequence and again in the boundary.
used_occurrences = {}


def resolve_sequence(names, description):
    resolved = []

    for name in names:
        matches = targets_by_name.get(name, [])
        occurrence = used_occurrences.get(name, 0)

        if occurrence >= len(matches):
            raise Exception(
                description
                + ": missing target occurrence "
                + str(occurrence + 1)
                + " for "
                + name
                + ". No robot movement has started."
            )

        resolved.append(matches[occurrence])
        used_occurrences[name] = occurrence + 1

    return resolved


# Resolve all target sequences before moving anything.
original_targets = resolve_sequence(
    original_names,
    "Original-side painting"
)

outline_targets = resolve_sequence(
    outline_names,
    "New-side outline"
)

boundary_targets = resolve_sequence(
    boundary_names,
    "Additional boundary"
)

# ------------------------------------------------------------
# VALIDATION REPORT
# ------------------------------------------------------------

print("\n============================================")
print("TARGET VALIDATION COMPLETE")
print("============================================")

print("Robot:", robot.Name())
print("Frame:", frame.Name())
print("Tool:", tool.Name())
print("Fixture:", fixture.Name())

print("Original-side targets:", len(original_targets))
print("New-side outline targets:", len(outline_targets))
print("Additional boundary targets:", len(boundary_targets))

print("\nOriginal-side sequence:")
for target in original_targets:
    print(" ->", target.Name())

print("\nNew-side outline sequence:")
for target in outline_targets:
    print(" ->", target.Name())

print("\nAdditional boundary sequence:")
for target in boundary_targets:
    print(" ->", target.Name())

# ------------------------------------------------------------
# CONFIGURE ROBOT
# ------------------------------------------------------------

robot.setPoseFrame(frame)
robot.setPoseTool(tool)
robot.setSpeed(ROBOT_SPEED)

# ------------------------------------------------------------
# PHASE 1: INITIAL HOME
# ------------------------------------------------------------

print("\n============================================")
print("PHASE 1: INITIAL HOME")
print("============================================")

robot.MoveJ(initial_home)

# ------------------------------------------------------------
# PHASE 2: ORIGINAL-SIDE PAINTING
# ------------------------------------------------------------

print("\n============================================")
print("PHASE 2: ORIGINAL-SIDE PAINTING")
print("============================================")

robot.MoveJ(original_targets[0])

for index, target in enumerate(original_targets[1:], start=2):
    print(
        "Original-side target",
        index,
        "of",
        len(original_targets),
        ":",
        target.Name()
    )

    robot.MoveL(target)

print("Original-side painting completed through Target 106.")

# ------------------------------------------------------------
# PHASE 3: HOME AFTER TARGET 106
# ------------------------------------------------------------

print("\n============================================")
print("PHASE 3: RETURN TO HOME")
print("============================================")

robot.MoveJ(home_after_106)

print("Robot reached Home after Target 106.")

# ------------------------------------------------------------
# PHASE 4: SLOW 180-DEGREE ROTATION
# ------------------------------------------------------------

print("\n============================================")
print("PHASE 4: ROTATE CAR BY 180 DEGREES")
print("============================================")

current_joints = fixture.Joints().list()

if len(current_joints) != 1:
    raise Exception(
        "Expected exactly one rotary joint. Found: "
        + str(current_joints)
    )

current_angle = current_joints[0]

# Choose the opposite orientation while keeping the target
# within the expected 0-360 degree range.
if current_angle + ROTATION_DEGREES <= 360.0:
    target_angle = current_angle + ROTATION_DEGREES
else:
    target_angle = current_angle - ROTATION_DEGREES

